// Characterization of the safe state per error class that had no test (#24 aim 6, step 1 of specs/plans/2026-11-02-reference-
// implementation-issue-24.md; the table is specs/design/monetcommon-safe-states.md). These tests pin what FB_MonetTelescopeControl
// does today on mock axes, with the line of the behaviour in a comment; they are not a specification. A test whose name ends in
// _Current pins a behaviour that differs from the target of the table (decision D4) and is flipped by the fix (step 7). The
// Roof_Request_* tests and No_Roof_Request_On_Focus_Error specify bCloseRoofRequest (step 7 PR 1, D9; no clock, no power-on). Every test
// owns a rig and runs over many PLC cycles (VAR_INST of the method, one Scan() per cycle). Failed checks are also noted in
// GVL_Diag.sFailures (printed by Run-Tests.ps1).
FUNCTION_BLOCK MonetSafeState_Tests EXTENDS TcUnit.FB_TestSuite
VAR
END_VAR

Hydraulics_Error_While_Tracking_Ramps_Then_Parks_In_Place();
Hydraulics_Pressure_Loss_While_Tracking_Parks_In_Place_Without_Ramp();
Cover_Error_At_PowerOn_Fails_And_Stays_Parked();
Cover_Error_During_Park_Ends_The_Park_Without_Closed();
Cover_Error_While_Tracking_Drives_To_Park();
Estop_During_Slew_Locks_Then_Parks_In_Place_After_The_Release();
Safety_Error_While_Tracking_Locks_Then_Parks_In_Place_When_It_Clears();
Power_Failure_During_Goto_Ramps_Then_Parks_In_Place();
Power_Failure_With_Pressure_Loss_Parks_In_Place_Without_Ramp();
Goto_Times_Out_Ramps_Then_Drives_To_Park();
Home_Times_Out_Ramps_Then_Drives_To_Park();
Clock_Invalid_Slew_Input_Is_Rejected();
Watchdog_Parks_And_Closes_The_Roof_In_One_Scan();
Invalid_Motion_Config_Is_Software_Error_32();
Roof_Request_On_Axis_Errors();
Roof_Request_On_Hydraulics_Error();
Roof_Request_On_Estop();
Roof_Request_On_Safety_Error();
Roof_Request_On_Power_Failure();
No_Roof_Request_On_Focus_Error();

// #24 step 7 PR 3 (D8, row hydraulics error; until 0.13.0 Hydraulics_Error_While_Tracking_Keeps_Tracking_Current): a hydraulics error
// with the pressure still there (brake open) is a telescope error (bHwError) and ramps first: in the scan of the error bStop is set
// (stop transaction, #96) and the axes stay enabled; every axis is sent its MC_Stop while still enabled (no 0x4257). After the stop
// has settled the emergency park queued behind it (bParkAfterStop) parks in place: axes disabled, brake closed, covers closed,
// hydraulics off, bIsParked and bParkedInPlace; READY_STATE -1.0 and bCloseRoofRequest while the error stays.
METHOD PRIVATE Hydraulics_Error_While_Tracking_Ramps_Then_Parks_In_Place
VAR_INST
	rig			: FB_MonetRig;
	nStep		: INT;
	nCycles		: UINT;
	nTracking	: UINT;
	sTest		: STRING(80);
	nEl0		: UINT;	// stop edges per axis before the error
	nAz0		: UINT;
	nDr0		: UINT;
	nExt0		: UINT;	// 0x4257 rejections of the three axes before the error
	nEdgesLast	: UINT;
	nEdgesNow	: UINT;
	nDisable0	: UINT;
	bSawStop	: BOOL;
	bStopOnDisabled	: BOOL;	// a stop edge came in a scan in which an axis was already disabled
END_VAR
TEST('Hydraulics_Error_While_Tracking_Ramps_Then_Parks_In_Place');
sTest := 'Hydraulics_Error_While_Tracking_Ramps_Then_Parks_In_Place: ';
IF nStep >= 90 THEN
	RETURN;
END_IF
rig.Scan();
nCycles := nCycles + 1;
CASE nStep OF
0:	// wait for the clock, then power on
	IF rig.ClockValid THEN
		rig.fbTel.Init();
		nStep := 10;
		nCycles := 0;
	ELSIF nCycles > 2000 THEN
		AssertTrue(Condition := FALSE, Message := 'the astronomical clock never became valid');
		F_Note(bFailed := TRUE, sText := CONCAT(sTest, 'the astronomical clock never became valid'));
		nStep := 99;
		TEST_FINISHED();
	END_IF
10:	// online: track a circumpolar target (always above the horizon, any RA)
	IF rig.Online THEN
		rig.fbTel.Track(fRightAscension := 0.0, fDeclination := -85.0);
		nStep := 20;
		nCycles := 0;
	ELSIF nCycles > 1500 THEN
		AssertTrue(Condition := FALSE, Message := 'the mock telescope did not reach READY_STATE 1.0');
		F_Note(bFailed := TRUE, sText := CONCAT(sTest, 'the mock telescope did not reach READY_STATE 1.0'));
		nStep := 99;
		TEST_FINISHED();
	END_IF
20:	// wait until all three axes have tracked for a few scans, then the hydraulics report an error (pressure still there)
	IF rig.fbAzim.Tracking AND rig.fbElev.Tracking AND rig.fbDero.Tracking THEN
		nTracking := nTracking + 1;
	ELSE
		nTracking := 0;
	END_IF
	IF nTracking >= 5 THEN
		nEl0 := rig.fbElev.nStopEdges;
		nAz0 := rig.fbAzim.nStopEdges;
		nDr0 := rig.fbDero.nStopEdges;
		nEdgesLast := nEl0 + nAz0 + nDr0;
		nExt0 := rig.fbElev.nExtErrors + rig.fbAzim.nExtErrors + rig.fbDero.nExtErrors;
		nDisable0 := rig.fbBrakeHyd.nDisableCalls;
		rig.fbBrakeHyd.InjectError();
		nStep := 30;
		nCycles := 0;
	ELSIF nCycles > 800 THEN
		AssertTrue(Condition := FALSE, Message := 'the telescope did not start tracking');
		F_Note(bFailed := TRUE, sText := CONCAT(sTest, 'the telescope did not start tracking'));
		nStep := 99;
		TEST_FINISHED();
	END_IF
30:	// ramp, then the park in place
	bSawStop := bSawStop OR rig.fbTel.bStopActive;
	nEdgesNow := rig.fbElev.nStopEdges + rig.fbAzim.nStopEdges + rig.fbDero.nStopEdges;
	IF nEdgesNow > nEdgesLast AND NOT (rig.fbElev.bEnable AND rig.fbAzim.bEnable AND rig.fbDero.bEnable) THEN
		bStopOnDisabled := TRUE;
	END_IF
	nEdgesLast := nEdgesNow;
	IF nCycles = 1 THEN	// the scan that saw the error
		AssertTrue(Condition := rig.fbTel.bStopActive AND rig.fbTel.bError, Message := 'the error stops the axes in its scan (bStop) and is a telescope error');
		F_Note(bFailed := NOT (rig.fbTel.bStopActive AND rig.fbTel.bError), sText := CONCAT(sTest, 'the error stops the axes in its scan (bStop) and is a telescope error'));
		AssertTrue(Condition := rig.fbElev.bEnable AND rig.fbAzim.bEnable AND rig.fbDero.bEnable, Message := 'the axes stay enabled for the ramp');
		F_Note(bFailed := NOT (rig.fbElev.bEnable AND rig.fbAzim.bEnable AND rig.fbDero.bEnable), sText := CONCAT(sTest, 'the axes stay enabled for the ramp'));
	END_IF
	IF rig.fbTel.bIsParked AND nCycles > 5 THEN
		AssertTrue(Condition := bSawStop, Message := 'the hydraulics error ramped (bStop)');
		F_Note(bFailed := NOT (bSawStop), sText := CONCAT(sTest, 'the hydraulics error ramped (bStop)'));
		AssertTrue(Condition := rig.fbElev.nStopEdges > nEl0 AND rig.fbAzim.nStopEdges > nAz0 AND rig.fbDero.nStopEdges > nDr0, Message := 'every axis was sent its MC_Stop');
		F_Note(bFailed := NOT (rig.fbElev.nStopEdges > nEl0 AND rig.fbAzim.nStopEdges > nAz0 AND rig.fbDero.nStopEdges > nDr0), sText := CONCAT(sTest, 'every axis was sent its MC_Stop'));
		AssertFalse(Condition := bStopOnDisabled, Message := 'the stops came before the disable');
		F_Note(bFailed := (bStopOnDisabled), sText := CONCAT(sTest, 'the stops came before the disable'));
		AssertTrue(Condition := rig.fbElev.nExtErrors + rig.fbAzim.nExtErrors + rig.fbDero.nExtErrors = nExt0, Message := 'no stop met the setpoint generator (0x4257)');
		F_Note(bFailed := NOT (rig.fbElev.nExtErrors + rig.fbAzim.nExtErrors + rig.fbDero.nExtErrors = nExt0), sText := CONCAT(sTest, 'no stop met the setpoint generator (0x4257)'));
		AssertTrue(Condition := rig.fbTel.bParkedInPlace AND NOT rig.fbTel.bParkActive, Message := 'the park ended in place');
		F_Note(bFailed := NOT (rig.fbTel.bParkedInPlace AND NOT rig.fbTel.bParkActive), sText := CONCAT(sTest, 'the park ended in place'));
		AssertFalse(Condition := rig.fbElev.bEnable OR rig.fbAzim.bEnable OR rig.fbDero.bEnable, Message := 'all three axes are disabled');
		F_Note(bFailed := (rig.fbElev.bEnable OR rig.fbAzim.bEnable OR rig.fbDero.bEnable), sText := CONCAT(sTest, 'all three axes are disabled'));
		AssertFalse(Condition := rig.fbBrakeHyd.BrakeOpen, Message := 'the brake is closed');
		F_Note(bFailed := (rig.fbBrakeHyd.BrakeOpen), sText := CONCAT(sTest, 'the brake is closed'));
		AssertTrue(Condition := rig.fbCovers.bClosed AND rig.fbCovers.nCloseCalls >= 1, Message := 'the covers are closed');
		F_Note(bFailed := NOT (rig.fbCovers.bClosed AND rig.fbCovers.nCloseCalls >= 1), sText := CONCAT(sTest, 'the covers are closed'));
		AssertTrue(Condition := rig.fbBrakeHyd.nDisableCalls > nDisable0, Message := 'the hydraulics are switched off');
		F_Note(bFailed := NOT (rig.fbBrakeHyd.nDisableCalls > nDisable0), sText := CONCAT(sTest, 'the hydraulics are switched off'));
		AssertFalse(Condition := rig.fbTel.bTrackActive OR rig.fbAzim.Tracking OR rig.fbElev.Tracking OR rig.fbDero.Tracking, Message := 'nothing tracks any more');
		F_Note(bFailed := (rig.fbTel.bTrackActive OR rig.fbAzim.Tracking OR rig.fbElev.Tracking OR rig.fbDero.Tracking), sText := CONCAT(sTest, 'nothing tracks any more'));
		AssertTrue(Condition := rig.fbTel.bError AND rig.fbTel.ReadyState = -1.0, Message := 'the error stays, READY_STATE -1.0');
		F_Note(bFailed := NOT (rig.fbTel.bError AND rig.fbTel.ReadyState = -1.0), sText := CONCAT(sTest, 'the error stays, READY_STATE -1.0'));
		AssertTrue(Condition := rig.fbTel.bCloseRoofRequest, Message := 'the roof close is requested');
		F_Note(bFailed := NOT (rig.fbTel.bCloseRoofRequest), sText := CONCAT(sTest, 'the roof close is requested'));
		nStep := 99;
		TEST_FINISHED();
	ELSIF nCycles > 800 THEN
		AssertTrue(Condition := FALSE, Message := 'the telescope did not park after the ramp');
		F_Note(bFailed := TRUE, sText := CONCAT(sTest, 'the telescope did not park after the ramp'));
		nStep := 99;
		TEST_FINISHED();
	END_IF
END_CASE
END_METHOD

// #24 step 7 PR 3 (D8, row hydraulics error): a hydraulics error with the oil pressure already gone (mock InjectPressureLoss: the
// brake is locked) cannot ramp, the brake lock is the stop: the axes are disabled in the scan of the error, as for an axis error,
// no MC_Stop is sent, and the emergency park parks in place (covers closed, hydraulics off, bIsParked, bParkedInPlace).
METHOD PRIVATE Hydraulics_Pressure_Loss_While_Tracking_Parks_In_Place_Without_Ramp
VAR_INST
	rig			: FB_MonetRig;
	nStep		: INT;
	nCycles		: UINT;
	nTracking	: UINT;
	sTest		: STRING(80);
	nEdges0		: UINT;	// stop edges of the three axes before the error
	nDisable0	: UINT;
	bSawStop	: BOOL;
END_VAR
TEST('Hydraulics_Pressure_Loss_While_Tracking_Parks_In_Place_Without_Ramp');
sTest := 'Hydraulics_Pressure_Loss_While_Tracking_Parks_In_Place_Without_Ramp: ';
IF nStep >= 90 THEN
	RETURN;
END_IF
rig.Scan();
nCycles := nCycles + 1;
CASE nStep OF
0:	// wait for the clock, then power on
	IF rig.ClockValid THEN
		rig.fbTel.Init();
		nStep := 10;
		nCycles := 0;
	ELSIF nCycles > 2000 THEN
		AssertTrue(Condition := FALSE, Message := 'the astronomical clock never became valid');
		F_Note(bFailed := TRUE, sText := CONCAT(sTest, 'the astronomical clock never became valid'));
		nStep := 99;
		TEST_FINISHED();
	END_IF
10:	// online: track a circumpolar target
	IF rig.Online THEN
		rig.fbTel.Track(fRightAscension := 0.0, fDeclination := -85.0);
		nStep := 20;
		nCycles := 0;
	ELSIF nCycles > 1500 THEN
		AssertTrue(Condition := FALSE, Message := 'the mock telescope did not reach READY_STATE 1.0');
		F_Note(bFailed := TRUE, sText := CONCAT(sTest, 'the mock telescope did not reach READY_STATE 1.0'));
		nStep := 99;
		TEST_FINISHED();
	END_IF
20:	// tracking: the hydraulics fail and the pressure is gone at once (the brake locks)
	IF rig.fbAzim.Tracking AND rig.fbElev.Tracking AND rig.fbDero.Tracking THEN
		nTracking := nTracking + 1;
	ELSE
		nTracking := 0;
	END_IF
	IF nTracking >= 5 THEN
		nEdges0 := rig.fbElev.nStopEdges + rig.fbAzim.nStopEdges + rig.fbDero.nStopEdges;
		nDisable0 := rig.fbBrakeHyd.nDisableCalls;
		rig.fbBrakeHyd.InjectPressureLoss();
		nStep := 30;
		nCycles := 0;
	ELSIF nCycles > 800 THEN
		AssertTrue(Condition := FALSE, Message := 'the telescope did not start tracking');
		F_Note(bFailed := TRUE, sText := CONCAT(sTest, 'the telescope did not start tracking'));
		nStep := 99;
		TEST_FINISHED();
	END_IF
30:
	bSawStop := bSawStop OR rig.fbTel.bStopActive;
	IF nCycles = 1 THEN	// the scan that saw the error
		AssertFalse(Condition := rig.fbElev.bEnable OR rig.fbAzim.bEnable OR rig.fbDero.bEnable, Message := 'the lock is the stop: disabled in the scan of the error');
		F_Note(bFailed := (rig.fbElev.bEnable OR rig.fbAzim.bEnable OR rig.fbDero.bEnable), sText := CONCAT(sTest, 'the lock is the stop: disabled in the scan of the error'));
	END_IF
	IF rig.fbTel.bIsParked AND nCycles > 5 THEN
		AssertFalse(Condition := bSawStop, Message := 'no ramp (bStop never set)');
		F_Note(bFailed := (bSawStop), sText := CONCAT(sTest, 'no ramp (bStop never set)'));
		AssertTrue(Condition := rig.fbElev.nStopEdges + rig.fbAzim.nStopEdges + rig.fbDero.nStopEdges = nEdges0, Message := 'no MC_Stop was sent');
		F_Note(bFailed := NOT (rig.fbElev.nStopEdges + rig.fbAzim.nStopEdges + rig.fbDero.nStopEdges = nEdges0), sText := CONCAT(sTest, 'no MC_Stop was sent'));
		AssertTrue(Condition := rig.fbTel.bParkedInPlace AND NOT rig.fbTel.bParkActive, Message := 'the park ended in place');
		F_Note(bFailed := NOT (rig.fbTel.bParkedInPlace AND NOT rig.fbTel.bParkActive), sText := CONCAT(sTest, 'the park ended in place'));
		AssertFalse(Condition := rig.fbBrakeHyd.BrakeOpen, Message := 'the brake is locked');
		F_Note(bFailed := (rig.fbBrakeHyd.BrakeOpen), sText := CONCAT(sTest, 'the brake is locked'));
		AssertTrue(Condition := rig.fbCovers.bClosed AND rig.fbCovers.nCloseCalls >= 1, Message := 'the covers are closed');
		F_Note(bFailed := NOT (rig.fbCovers.bClosed AND rig.fbCovers.nCloseCalls >= 1), sText := CONCAT(sTest, 'the covers are closed'));
		AssertTrue(Condition := rig.fbBrakeHyd.nDisableCalls > nDisable0, Message := 'the hydraulics are switched off');
		F_Note(bFailed := NOT (rig.fbBrakeHyd.nDisableCalls > nDisable0), sText := CONCAT(sTest, 'the hydraulics are switched off'));
		AssertTrue(Condition := rig.fbTel.bError AND rig.fbTel.ReadyState = -1.0, Message := 'the error stays, READY_STATE -1.0');
		F_Note(bFailed := NOT (rig.fbTel.bError AND rig.fbTel.ReadyState = -1.0), sText := CONCAT(sTest, 'the error stays, READY_STATE -1.0'));
		AssertTrue(Condition := rig.fbTel.bCloseRoofRequest, Message := 'the roof close is requested');
		F_Note(bFailed := NOT (rig.fbTel.bCloseRoofRequest), sText := CONCAT(sTest, 'the roof close is requested'));
		nStep := 99;
		TEST_FINISHED();
	ELSIF nCycles > 800 THEN
		AssertTrue(Condition := FALSE, Message := 'the emergency park did not finish');
		F_Note(bFailed := TRUE, sText := CONCAT(sTest, 'the emergency park did not finish'));
		nStep := 99;
		TEST_FINISHED();
	END_IF
END_CASE
END_METHOD

// #24 step 7 PR 4 (row cover error; until 0.13.x Cover_Error_At_PowerOn_Waits_In_Stage_0_Current, where the power-on waited in
// stage 0 for fbCovers.Opened until the 12 h command timeout, with bIsParked already FALSE). A cover error on a parked telescope
// starts no park. A power-on with the cover error fails in its first scan, before the cover command of stage 0 (_PowerOn checks,
// bPowerFailure): nothing opens, no axis is enabled, the telescope stays parked, READY_STATE -1.0, no telescope error, no roof
// close request (D9). Reset path: the cover reset (HalfBROT Reset(), MAIN reset button), then power=1 goes online.
METHOD PRIVATE Cover_Error_At_PowerOn_Fails_And_Stays_Parked
VAR_INST
	rig			: FB_MonetRig;
	nStep		: INT;
	nCycles		: UINT;
	sTest		: STRING(80);
END_VAR
TEST('Cover_Error_At_PowerOn_Fails_And_Stays_Parked');
sTest := 'Cover_Error_At_PowerOn_Fails_And_Stays_Parked: ';
IF nStep >= 90 THEN
	RETURN;
END_IF
rig.Scan();
nCycles := nCycles + 1;
CASE nStep OF
0:	// wait for the clock; the covers of the parked telescope report an error
	IF rig.ClockValid THEN
		rig.fbCovers.InjectError();
		nStep := 5;
		nCycles := 0;
	ELSIF nCycles > 2000 THEN
		AssertTrue(Condition := FALSE, Message := 'the astronomical clock never became valid');
		F_Note(bFailed := TRUE, sText := CONCAT(sTest, 'the astronomical clock never became valid'));
		nStep := 99;
		TEST_FINISHED();
	END_IF
5:	// parked: nothing happens; then power on
	IF nCycles >= 10 THEN
		AssertTrue(Condition := rig.fbTel.bIsParked AND NOT rig.fbTel.bParkActive AND NOT rig.fbTel.bError, Message := 'a cover error on a parked telescope starts no park and is no telescope error');
		F_Note(bFailed := NOT (rig.fbTel.bIsParked AND NOT rig.fbTel.bParkActive AND NOT rig.fbTel.bError), sText := CONCAT(sTest, 'a cover error on a parked telescope starts no park and is no telescope error'));
		rig.fbTel.Init();
		nStep := 10;
		nCycles := 0;
	END_IF
10:	// the power-on fails in its first scan
	IF nCycles >= 10 THEN
		AssertFalse(Condition := rig.fbTel.bPowerActive OR rig.fbTel.fbStartup.Initializing, Message := 'the power-on is over');
		F_Note(bFailed := (rig.fbTel.bPowerActive OR rig.fbTel.fbStartup.Initializing), sText := CONCAT(sTest, 'the power-on is over'));
		AssertTrue(Condition := rig.fbTel.bPowerFailure AND rig.fbTel.ReadyState = -1.0, Message := 'power-on failure, READY_STATE -1.0');
		F_Note(bFailed := NOT (rig.fbTel.bPowerFailure AND rig.fbTel.ReadyState = -1.0), sText := CONCAT(sTest, 'power-on failure, READY_STATE -1.0'));
		AssertTrue(Condition := rig.fbCovers.nOpenCalls = 0 AND NOT rig.fbCovers.bOpened, Message := 'the covers were not commanded');
		F_Note(bFailed := NOT (rig.fbCovers.nOpenCalls = 0 AND NOT rig.fbCovers.bOpened), sText := CONCAT(sTest, 'the covers were not commanded'));
		AssertFalse(Condition := rig.fbElev.bEnable OR rig.fbAzim.bEnable OR rig.fbDero.bEnable, Message := 'no axis was enabled');
		F_Note(bFailed := (rig.fbElev.bEnable OR rig.fbAzim.bEnable OR rig.fbDero.bEnable), sText := CONCAT(sTest, 'no axis was enabled'));
		AssertTrue(Condition := rig.fbTel.bIsParked, Message := 'the telescope stays parked');
		F_Note(bFailed := NOT (rig.fbTel.bIsParked), sText := CONCAT(sTest, 'the telescope stays parked'));
		AssertFalse(Condition := rig.fbTel.bError, Message := 'a cover error is not a telescope error');
		F_Note(bFailed := (rig.fbTel.bError), sText := CONCAT(sTest, 'a cover error is not a telescope error'));
		AssertFalse(Condition := rig.fbTel.bCloseRoofRequest, Message := 'no roof close request for a cover error');
		F_Note(bFailed := (rig.fbTel.bCloseRoofRequest), sText := CONCAT(sTest, 'no roof close request for a cover error'));
		rig.fbCovers.Reset();	// MAIN reset button
		nStep := 20;
		nCycles := 0;
	END_IF
20:
	IF nCycles >= 3 THEN
		rig.fbTel.Init();
		nStep := 30;
		nCycles := 0;
	END_IF
30:	// power=1 after the cover reset: online
	IF rig.Online THEN
		AssertTrue(Condition := rig.fbCovers.bOpened AND NOT rig.fbTel.bPowerFailure, Message := 'online after the cover reset and power=1');
		F_Note(bFailed := NOT (rig.fbCovers.bOpened AND NOT rig.fbTel.bPowerFailure), sText := CONCAT(sTest, 'online after the cover reset and power=1'));
		nStep := 99;
		TEST_FINISHED();
	ELSIF nCycles > 1500 THEN
		AssertTrue(Condition := FALSE, Message := 'not online after the cover reset and power=1');
		F_Note(bFailed := TRUE, sText := CONCAT(sTest, 'not online after the cover reset and power=1'));
		nStep := 99;
		TEST_FINISHED();
	END_IF
END_CASE
END_METHOD

// #24 step 7 PR 4 (row cover error; until 0.13.x Cover_Error_Holds_The_Park_Before_Parked_Current, where the park waited in stage
// secure for fbCovers.Closed for ever: bPark held, READY_STATE 0.3, never bIsParked). A cover error during the drive to the park
// position: the park goes on (no telescope error, the drives are controllable), reaches the park position, disables the axes, the
// brake closes, the hydraulics go off, and the park ends without Closed: bIsParked, not in place, software error 16#21 (READY_STATE
// -1.0), no roof close request (D9).
METHOD PRIVATE Cover_Error_During_Park_Ends_The_Park_Without_Closed
VAR_INST
	rig			: FB_MonetRig;
	nStep		: INT;
	nCycles		: UINT;
	sTest		: STRING(80);
	nDisable0	: UINT;
	bSawError	: BOOL;	// bError before the park ended
END_VAR
TEST('Cover_Error_During_Park_Ends_The_Park_Without_Closed');
sTest := 'Cover_Error_During_Park_Ends_The_Park_Without_Closed: ';
IF nStep >= 90 THEN
	RETURN;
END_IF
rig.Scan();
nCycles := nCycles + 1;
CASE nStep OF
0:	// wait for the clock, then power on
	IF rig.ClockValid THEN
		rig.fbTel.Init();
		nStep := 10;
		nCycles := 0;
	ELSIF nCycles > 2000 THEN
		AssertTrue(Condition := FALSE, Message := 'the astronomical clock never became valid');
		F_Note(bFailed := TRUE, sText := CONCAT(sTest, 'the astronomical clock never became valid'));
		nStep := 99;
		TEST_FINISHED();
	END_IF
10:	// online: slow axes, park
	IF rig.Online THEN
		rig.SetMoveScans(nScans := 300);
		nDisable0 := rig.fbBrakeHyd.nDisableCalls;
		rig.fbTel.Park();
		nStep := 20;
		nCycles := 0;
	ELSIF nCycles > 1500 THEN
		AssertTrue(Condition := FALSE, Message := 'the mock telescope did not reach READY_STATE 1.0');
		F_Note(bFailed := TRUE, sText := CONCAT(sTest, 'the mock telescope did not reach READY_STATE 1.0'));
		nStep := 99;
		TEST_FINISHED();
	END_IF
20:	// the park drives: the covers report an error
	IF rig.fbElev.MoveAxis AND rig.fbAzim.MoveAxis AND rig.fbDero.MoveAxis AND nCycles > 5 THEN
		rig.fbCovers.InjectError();
		nStep := 30;
		nCycles := 0;
	ELSIF nCycles > 300 THEN
		AssertTrue(Condition := FALSE, Message := 'the park did not start the axis moves');
		F_Note(bFailed := TRUE, sText := CONCAT(sTest, 'the park did not start the axis moves'));
		nStep := 99;
		TEST_FINISHED();
	END_IF
30:	// the park goes on and ends
	IF rig.fbTel.bIsParked THEN
		AssertFalse(Condition := bSawError, Message := 'no telescope error during the drive');
		F_Note(bFailed := (bSawError), sText := CONCAT(sTest, 'no telescope error during the drive'));
		AssertFalse(Condition := rig.fbTel.bParkActive OR rig.fbTel.bParkedInPlace, Message := 'the park is over, not in place');
		F_Note(bFailed := (rig.fbTel.bParkActive OR rig.fbTel.bParkedInPlace), sText := CONCAT(sTest, 'the park is over, not in place'));
		AssertTrue(Condition := ABS(rig.fbElev.fActualPosition - 60.0) < 0.001 AND ABS(rig.fbAzim.fActualPosition - 175.0) < 0.001, Message := 'at the park position');
		F_Note(bFailed := NOT (ABS(rig.fbElev.fActualPosition - 60.0) < 0.001 AND ABS(rig.fbAzim.fActualPosition - 175.0) < 0.001), sText := CONCAT(sTest, 'at the park position'));
		AssertFalse(Condition := rig.fbElev.bEnable OR rig.fbAzim.bEnable OR rig.fbDero.bEnable, Message := 'all three axes are disabled');
		F_Note(bFailed := (rig.fbElev.bEnable OR rig.fbAzim.bEnable OR rig.fbDero.bEnable), sText := CONCAT(sTest, 'all three axes are disabled'));
		AssertFalse(Condition := rig.fbBrakeHyd.BrakeOpen, Message := 'the brake is closed');
		F_Note(bFailed := (rig.fbBrakeHyd.BrakeOpen), sText := CONCAT(sTest, 'the brake is closed'));
		AssertTrue(Condition := rig.fbBrakeHyd.nDisableCalls > nDisable0, Message := 'the hydraulics are switched off');
		F_Note(bFailed := NOT (rig.fbBrakeHyd.nDisableCalls > nDisable0), sText := CONCAT(sTest, 'the hydraulics are switched off'));
		AssertTrue(Condition := rig.fbCovers.nCloseCalls >= 1 AND NOT rig.fbCovers.bClosed, Message := 'the covers were commanded closed and did not move');
		F_Note(bFailed := NOT (rig.fbCovers.nCloseCalls >= 1 AND NOT rig.fbCovers.bClosed), sText := CONCAT(sTest, 'the covers were commanded closed and did not move'));
		AssertTrue(Condition := rig.fbTel.bError AND rig.fbTel.nErrorID = 16#21 AND rig.fbTel.ReadyState = -1.0, Message := 'software error 16#21, READY_STATE -1.0');
		F_Note(bFailed := NOT (rig.fbTel.bError AND rig.fbTel.nErrorID = 16#21 AND rig.fbTel.ReadyState = -1.0), sText := CONCAT(sTest, 'software error 16#21, READY_STATE -1.0'));
		AssertFalse(Condition := rig.fbTel.bCloseRoofRequest, Message := 'no roof close request for a cover error');
		F_Note(bFailed := (rig.fbTel.bCloseRoofRequest), sText := CONCAT(sTest, 'no roof close request for a cover error'));
		nStep := 99;
		TEST_FINISHED();
	ELSIF nCycles > 1500 THEN
		AssertTrue(Condition := FALSE, Message := 'the park did not end (it waits for the covers)');
		F_Note(bFailed := TRUE, sText := CONCAT(sTest, 'the park did not end (it waits for the covers)'));
		nStep := 99;
		TEST_FINISHED();
	END_IF
	bSawError := bSawError OR rig.fbTel.bError;	// after the check: 16#21 is raised in the scan that sets bIsParked
END_CASE
END_METHOD

// #24 step 7 PR 4 (row cover error, target "ramp; drive to park"): a cover error while tracking is no telescope error (the drives are
// controllable) and starts a normal park in its scan (Park(), the routing of an external park: the track is dropped, the axes stay
// enabled and drive to the park position). The park ends without Closed: bIsParked, not in place, hydraulics off, software error
// 16#21, no roof close request (D9).
METHOD PRIVATE Cover_Error_While_Tracking_Drives_To_Park
VAR_INST
	rig			: FB_MonetRig;
	nStep		: INT;
	nCycles		: UINT;
	nTracking	: UINT;
	sTest		: STRING(80);
	nDisable0	: UINT;
END_VAR
TEST('Cover_Error_While_Tracking_Drives_To_Park');
sTest := 'Cover_Error_While_Tracking_Drives_To_Park: ';
IF nStep >= 90 THEN
	RETURN;
END_IF
rig.Scan();
nCycles := nCycles + 1;
CASE nStep OF
0:	// wait for the clock, then power on
	IF rig.ClockValid THEN
		rig.fbTel.Init();
		nStep := 10;
		nCycles := 0;
	ELSIF nCycles > 2000 THEN
		AssertTrue(Condition := FALSE, Message := 'the astronomical clock never became valid');
		F_Note(bFailed := TRUE, sText := CONCAT(sTest, 'the astronomical clock never became valid'));
		nStep := 99;
		TEST_FINISHED();
	END_IF
10:	// online: track a circumpolar target
	IF rig.Online THEN
		rig.fbTel.Track(fRightAscension := 0.0, fDeclination := -85.0);
		nStep := 20;
		nCycles := 0;
	ELSIF nCycles > 1500 THEN
		AssertTrue(Condition := FALSE, Message := 'the mock telescope did not reach READY_STATE 1.0');
		F_Note(bFailed := TRUE, sText := CONCAT(sTest, 'the mock telescope did not reach READY_STATE 1.0'));
		nStep := 99;
		TEST_FINISHED();
	END_IF
20:	// tracking: the covers report an error
	IF rig.fbAzim.Tracking AND rig.fbElev.Tracking AND rig.fbDero.Tracking THEN
		nTracking := nTracking + 1;
	ELSE
		nTracking := 0;
	END_IF
	IF nTracking >= 5 THEN
		nDisable0 := rig.fbBrakeHyd.nDisableCalls;
		rig.fbCovers.InjectError();
		nStep := 30;
		nCycles := 0;
	ELSIF nCycles > 800 THEN
		AssertTrue(Condition := FALSE, Message := 'the telescope did not start tracking');
		F_Note(bFailed := TRUE, sText := CONCAT(sTest, 'the telescope did not start tracking'));
		nStep := 99;
		TEST_FINISHED();
	END_IF
30:
	IF nCycles = 1 THEN	// the scan that saw the error
		AssertTrue(Condition := rig.fbTel.bParkActive AND NOT rig.fbTel.bTrackActive, Message := 'the park is requested in the scan of the error, the track is dropped');
		F_Note(bFailed := NOT (rig.fbTel.bParkActive AND NOT rig.fbTel.bTrackActive), sText := CONCAT(sTest, 'the park is requested in the scan of the error, the track is dropped'));
		AssertTrue(Condition := NOT rig.fbTel.bError AND rig.fbElev.bEnable AND rig.fbAzim.bEnable AND rig.fbDero.bEnable, Message := 'no telescope error, the axes stay enabled');
		F_Note(bFailed := NOT (NOT rig.fbTel.bError AND rig.fbElev.bEnable AND rig.fbAzim.bEnable AND rig.fbDero.bEnable), sText := CONCAT(sTest, 'no telescope error, the axes stay enabled'));
	END_IF
	IF rig.fbTel.bIsParked AND nCycles > 5 THEN
		AssertFalse(Condition := rig.fbTel.bParkActive OR rig.fbTel.bParkedInPlace, Message := 'the park is over, not in place');
		F_Note(bFailed := (rig.fbTel.bParkActive OR rig.fbTel.bParkedInPlace), sText := CONCAT(sTest, 'the park is over, not in place'));
		AssertTrue(Condition := ABS(rig.fbElev.fActualPosition - 60.0) < 0.001 AND ABS(rig.fbAzim.fActualPosition - 175.0) < 0.001, Message := 'at the park position');
		F_Note(bFailed := NOT (ABS(rig.fbElev.fActualPosition - 60.0) < 0.001 AND ABS(rig.fbAzim.fActualPosition - 175.0) < 0.001), sText := CONCAT(sTest, 'at the park position'));
		AssertFalse(Condition := rig.fbTel.bTrackActive OR rig.fbAzim.Tracking OR rig.fbElev.Tracking OR rig.fbDero.Tracking, Message := 'nothing tracks any more');
		F_Note(bFailed := (rig.fbTel.bTrackActive OR rig.fbAzim.Tracking OR rig.fbElev.Tracking OR rig.fbDero.Tracking), sText := CONCAT(sTest, 'nothing tracks any more'));
		AssertFalse(Condition := rig.fbElev.bEnable OR rig.fbAzim.bEnable OR rig.fbDero.bEnable OR rig.fbBrakeHyd.BrakeOpen, Message := 'axes disabled, brake closed');
		F_Note(bFailed := (rig.fbElev.bEnable OR rig.fbAzim.bEnable OR rig.fbDero.bEnable OR rig.fbBrakeHyd.BrakeOpen), sText := CONCAT(sTest, 'axes disabled, brake closed'));
		AssertTrue(Condition := rig.fbBrakeHyd.nDisableCalls > nDisable0, Message := 'the hydraulics are switched off');
		F_Note(bFailed := NOT (rig.fbBrakeHyd.nDisableCalls > nDisable0), sText := CONCAT(sTest, 'the hydraulics are switched off'));
		AssertFalse(Condition := rig.fbCovers.bClosed, Message := 'the covers did not move');
		F_Note(bFailed := (rig.fbCovers.bClosed), sText := CONCAT(sTest, 'the covers did not move'));
		AssertTrue(Condition := rig.fbTel.nErrorID = 16#21 AND rig.fbTel.ReadyState = -1.0, Message := 'software error 16#21, READY_STATE -1.0');
		F_Note(bFailed := NOT (rig.fbTel.nErrorID = 16#21 AND rig.fbTel.ReadyState = -1.0), sText := CONCAT(sTest, 'software error 16#21, READY_STATE -1.0'));
		AssertFalse(Condition := rig.fbTel.bCloseRoofRequest, Message := 'no roof close request for a cover error');
		F_Note(bFailed := (rig.fbTel.bCloseRoofRequest), sText := CONCAT(sTest, 'no roof close request for a cover error'));
		nStep := 99;
		TEST_FINISHED();
	ELSIF nCycles > 1500 THEN
		AssertTrue(Condition := FALSE, Message := 'the park did not end');
		F_Note(bFailed := TRUE, sText := CONCAT(sTest, 'the park did not end'));
		nStep := 99;
		TEST_FINISHED();
	END_IF
END_CASE
END_METHOD

// #24 step 7 PR 6 (D8, row E-stop; until 0.13.0 Estop_During_Slew_Disables_The_Axes_Without_Park_Current): the E-stop under a slew
// is a lock stop: in its scan the three axes are disabled and the hydraulics switched off (the brake locks), no stop transaction
// (no bStop, no MC_Stop), the slew ends. During the E-stop nothing parks and the covers are not commanded (they may hang on the
// same circuit), also not after a reset (the MAIN reset button that starts the safety reset); READY_STATE -1.0, not bError. After
// the release (E-stop gone, safety reset done) the held park runs in place: covers closed, hydraulics off, bIsParked,
// bParkedInPlace; the roof request stays until a reset; then power=1 is online again. The mock axis keeps its move when it is
// disabled (STO is not modelled), so the test ends the mock move (SetMoveScans) before the release.
METHOD PRIVATE Estop_During_Slew_Locks_Then_Parks_In_Place_After_The_Release
VAR_INST
	rig			: FB_MonetRig;
	nStep		: INT;
	nCycles		: UINT;
	sTest		: STRING(80);
	nDisable0	: UINT;	// hydraulics-off writes before the E-stop
	nDisable1	: UINT;	// ... before the release
	nEdges0		: UINT;	// MC_Stop requests of the three axes before the E-stop
	bSawStop	: BOOL;
END_VAR
TEST('Estop_During_Slew_Locks_Then_Parks_In_Place_After_The_Release');
sTest := 'Estop_During_Slew_Locks_Then_Parks_In_Place_After_The_Release: ';
IF nStep >= 90 THEN
	RETURN;
END_IF
rig.Scan();
nCycles := nCycles + 1;
CASE nStep OF
0:	// wait for the clock, then power on
	IF rig.ClockValid THEN
		rig.fbTel.Init();
		nStep := 10;
		nCycles := 0;
	ELSIF nCycles > 2000 THEN
		AssertTrue(Condition := FALSE, Message := 'the astronomical clock never became valid');
		F_Note(bFailed := TRUE, sText := CONCAT(sTest, 'the astronomical clock never became valid'));
		nStep := 99;
		TEST_FINISHED();
	END_IF
10:	// online: slow axes, slew
	IF rig.Online THEN
		rig.SetMoveScans(nScans := 3000);
		rig.fbTel.Slew(fAzimuth := 180.0, fAltitude := 45.0);
		nStep := 20;
		nCycles := 0;
	ELSIF nCycles > 1500 THEN
		AssertTrue(Condition := FALSE, Message := 'the mock telescope did not reach READY_STATE 1.0');
		F_Note(bFailed := TRUE, sText := CONCAT(sTest, 'the mock telescope did not reach READY_STATE 1.0'));
		nStep := 99;
		TEST_FINISHED();
	END_IF
20:
	IF rig.fbElev.MoveAxis AND rig.fbAzim.MoveAxis AND rig.fbDero.MoveAxis THEN
		nStep := 30;
		nCycles := 0;
	ELSIF nCycles > 300 THEN
		AssertTrue(Condition := FALSE, Message := 'the slew did not start the axis moves');
		F_Note(bFailed := TRUE, sText := CONCAT(sTest, 'the slew did not start the axis moves'));
		nStep := 99;
		TEST_FINISHED();
	END_IF
30:	// the axes move: the E-stop is pressed
	IF nCycles >= 5 THEN
		nDisable0 := rig.fbBrakeHyd.nDisableCalls;
		nEdges0 := rig.fbElev.nStopEdges + rig.fbAzim.nStopEdges + rig.fbDero.nStopEdges;
		rig.SetEstop(TRUE);
		nStep := 40;
		nCycles := 0;
	END_IF
40:	// the lock is the stop; the park is held while the E-stop is pressed
	bSawStop := bSawStop OR rig.fbTel.bStopActive;
	IF nCycles = 1 THEN	// the scan that saw the E-stop
		AssertFalse(Condition := rig.fbElev.bEnable OR rig.fbAzim.bEnable OR rig.fbDero.bEnable, Message := 'the axes are disabled in the scan of the E-stop');
		F_Note(bFailed := (rig.fbElev.bEnable OR rig.fbAzim.bEnable OR rig.fbDero.bEnable), sText := CONCAT(sTest, 'the axes are disabled in the scan of the E-stop'));
		AssertTrue(Condition := rig.fbBrakeHyd.nDisableCalls > nDisable0, Message := 'the hydraulics go off in the scan of the E-stop');
		F_Note(bFailed := NOT (rig.fbBrakeHyd.nDisableCalls > nDisable0), sText := CONCAT(sTest, 'the hydraulics go off in the scan of the E-stop'));
		AssertTrue(Condition := rig.fbCovers.nStopCalls >= 1, Message := 'the covers get Stop() in the scan of the E-stop (not on the E-stop circuit)');
		F_Note(bFailed := NOT (rig.fbCovers.nStopCalls >= 1), sText := CONCAT(sTest, 'the covers get Stop() in the scan of the E-stop (not on the E-stop circuit)'));
	END_IF
	IF nCycles >= 60 THEN
		AssertFalse(Condition := rig.fbElev.bEnable OR rig.fbAzim.bEnable OR rig.fbDero.bEnable, Message := 'the three axes are disabled');
		F_Note(bFailed := (rig.fbElev.bEnable OR rig.fbAzim.bEnable OR rig.fbDero.bEnable), sText := CONCAT(sTest, 'the three axes are disabled'));
		AssertFalse(Condition := rig.fbBrakeHyd.BrakeOpen, Message := 'the brake is closed');
		F_Note(bFailed := (rig.fbBrakeHyd.BrakeOpen), sText := CONCAT(sTest, 'the brake is closed'));
		AssertFalse(Condition := bSawStop, Message := 'no ramp (bStop never set)');
		F_Note(bFailed := (bSawStop), sText := CONCAT(sTest, 'no ramp (bStop never set)'));
		AssertTrue(Condition := rig.fbElev.nStopEdges + rig.fbAzim.nStopEdges + rig.fbDero.nStopEdges = nEdges0, Message := 'no MC_Stop was sent');
		F_Note(bFailed := NOT (rig.fbElev.nStopEdges + rig.fbAzim.nStopEdges + rig.fbDero.nStopEdges = nEdges0), sText := CONCAT(sTest, 'no MC_Stop was sent'));
		AssertFalse(Condition := rig.fbTel.bSlewActive, Message := 'the slew has ended');
		F_Note(bFailed := (rig.fbTel.bSlewActive), sText := CONCAT(sTest, 'the slew has ended'));
		AssertFalse(Condition := rig.fbTel.bParkActive OR rig.fbTel.bIsParked, Message := 'no park during the E-stop');
		F_Note(bFailed := (rig.fbTel.bParkActive OR rig.fbTel.bIsParked), sText := CONCAT(sTest, 'no park during the E-stop'));
		AssertTrue(Condition := rig.fbCovers.nCloseCalls = 0, Message := 'the covers are not commanded during the E-stop');
		F_Note(bFailed := NOT (rig.fbCovers.nCloseCalls = 0), sText := CONCAT(sTest, 'the covers are not commanded during the E-stop'));
		AssertFalse(Condition := rig.fbTel.bError, Message := 'the E-stop is not bError');
		F_Note(bFailed := (rig.fbTel.bError), sText := CONCAT(sTest, 'the E-stop is not bError'));
		AssertTrue(Condition := rig.fbTel.ReadyState = -1.0, Message := 'READY_STATE is -1.0');
		F_Note(bFailed := NOT (rig.fbTel.ReadyState = -1.0), sText := CONCAT(sTest, 'READY_STATE is -1.0'));
		rig.SetMoveScans(nScans := 60);	// STO is not modelled: end the move the disabled mock axes still run
		rig.fbTel.Reset();	// the MAIN reset button during the E-stop (starts the safety reset)
		nStep := 50;
		nCycles := 0;
	END_IF
50:	// a reset during the E-stop does not start the park
	bSawStop := bSawStop OR rig.fbTel.bStopActive;
	IF nCycles >= 10 THEN
		AssertTrue(Condition := NOT (rig.fbTel.bParkActive OR rig.fbTel.bIsParked) AND rig.fbCovers.nCloseCalls = 0, Message := 'a reset during the E-stop does not start the park');
		F_Note(bFailed := NOT (NOT (rig.fbTel.bParkActive OR rig.fbTel.bIsParked) AND rig.fbCovers.nCloseCalls = 0), sText := CONCAT(sTest, 'a reset during the E-stop does not start the park'));
		nDisable1 := rig.fbBrakeHyd.nDisableCalls;
		rig.SetEstop(FALSE);	// released, safety reset done
		nStep := 60;
		nCycles := 0;
	END_IF
60:	// after the release: the park in place
	bSawStop := bSawStop OR rig.fbTel.bStopActive;
	IF rig.fbTel.bIsParked AND nCycles > 5 THEN
		AssertTrue(Condition := rig.fbTel.bParkedInPlace AND NOT rig.fbTel.bParkActive, Message := 'the park after the release ended in place');
		F_Note(bFailed := NOT (rig.fbTel.bParkedInPlace AND NOT rig.fbTel.bParkActive), sText := CONCAT(sTest, 'the park after the release ended in place'));
		AssertTrue(Condition := rig.fbCovers.bClosed AND rig.fbCovers.nCloseCalls >= 1, Message := 'the covers are closed after the release');
		F_Note(bFailed := NOT (rig.fbCovers.bClosed AND rig.fbCovers.nCloseCalls >= 1), sText := CONCAT(sTest, 'the covers are closed after the release'));
		AssertTrue(Condition := rig.fbBrakeHyd.nDisableCalls > nDisable1, Message := 'the park switches the hydraulics off');
		F_Note(bFailed := NOT (rig.fbBrakeHyd.nDisableCalls > nDisable1), sText := CONCAT(sTest, 'the park switches the hydraulics off'));
		AssertFalse(Condition := rig.fbElev.bEnable OR rig.fbAzim.bEnable OR rig.fbDero.bEnable OR rig.fbBrakeHyd.BrakeOpen, Message := 'axes disabled, brake closed');
		F_Note(bFailed := (rig.fbElev.bEnable OR rig.fbAzim.bEnable OR rig.fbDero.bEnable OR rig.fbBrakeHyd.BrakeOpen), sText := CONCAT(sTest, 'axes disabled, brake closed'));
		AssertFalse(Condition := bSawStop, Message := 'no stop at all');
		F_Note(bFailed := (bSawStop), sText := CONCAT(sTest, 'no stop at all'));
		AssertTrue(Condition := rig.fbTel.bCloseRoofRequest, Message := 'the roof request stays latched');
		F_Note(bFailed := NOT (rig.fbTel.bCloseRoofRequest), sText := CONCAT(sTest, 'the roof request stays latched'));
		rig.fbTel.Reset();
		nStep := 70;
		nCycles := 0;
	ELSIF nCycles > 600 THEN
		AssertTrue(Condition := FALSE, Message := 'the park after the release did not finish');
		F_Note(bFailed := TRUE, sText := CONCAT(sTest, 'the park after the release did not finish'));
		nStep := 99;
		TEST_FINISHED();
	END_IF
70:
	IF nCycles >= 10 THEN
		AssertFalse(Condition := rig.fbTel.bCloseRoofRequest, Message := 'the reset after the release clears the roof request');
		F_Note(bFailed := (rig.fbTel.bCloseRoofRequest), sText := CONCAT(sTest, 'the reset after the release clears the roof request'));
		rig.fbTel.Init();
		nStep := 80;
		nCycles := 0;
	END_IF
80:	// power=1: online again
	IF rig.Online THEN
		AssertTrue(Condition := TRUE, Message := 'online again after the release, the reset and power=1');
		nStep := 99;
		TEST_FINISHED();
	ELSIF nCycles > 1500 THEN
		AssertTrue(Condition := FALSE, Message := 'not online again after the release, the reset and power=1');
		F_Note(bFailed := TRUE, sText := CONCAT(sTest, 'not online again after the release, the reset and power=1'));
		nStep := 99;
		TEST_FINISHED();
	END_IF
END_CASE
END_METHOD

// #24 step 7 PR 6 (D8, row safety error; until 0.13.0 a safety error without E-stop only acted on the brake in the Wake&Shake window):
// a safety error (SafetyHandling.error, no E-stop) under tracking is handled as the E-stop: in its scan the axes are disabled and the
// hydraulics switched off (the lock is the stop, no bStop, no MC_Stop), tracking ends; nothing parks and the covers are not
// commanded while it is there (it is not bError); the roof close is requested. When it is gone the held park runs in place.
METHOD PRIVATE Safety_Error_While_Tracking_Locks_Then_Parks_In_Place_When_It_Clears
VAR_INST
	rig			: FB_MonetRig;
	nStep		: INT;
	nCycles		: UINT;
	nTracking	: UINT;
	sTest		: STRING(80);
	nDisable0	: UINT;	// hydraulics-off writes before the safety error
	nDisable1	: UINT;	// ... before it clears
	nEdges0		: UINT;	// MC_Stop requests of the three axes before the safety error
	bSawStop	: BOOL;
END_VAR
TEST('Safety_Error_While_Tracking_Locks_Then_Parks_In_Place_When_It_Clears');
sTest := 'Safety_Error_While_Tracking_Locks_Then_Parks_In_Place_When_It_Clears: ';
IF nStep >= 90 THEN
	RETURN;
END_IF
rig.Scan();
nCycles := nCycles + 1;
CASE nStep OF
0:	// wait for the clock, then power on
	IF rig.ClockValid THEN
		rig.fbTel.Init();
		nStep := 10;
		nCycles := 0;
	ELSIF nCycles > 2000 THEN
		AssertTrue(Condition := FALSE, Message := 'the astronomical clock never became valid');
		F_Note(bFailed := TRUE, sText := CONCAT(sTest, 'the astronomical clock never became valid'));
		nStep := 99;
		TEST_FINISHED();
	END_IF
10:	// online: track a circumpolar target
	IF rig.Online THEN
		rig.fbTel.Track(fRightAscension := 0.0, fDeclination := -85.0);
		nStep := 20;
		nCycles := 0;
	ELSIF nCycles > 1500 THEN
		AssertTrue(Condition := FALSE, Message := 'the mock telescope did not reach READY_STATE 1.0');
		F_Note(bFailed := TRUE, sText := CONCAT(sTest, 'the mock telescope did not reach READY_STATE 1.0'));
		nStep := 99;
		TEST_FINISHED();
	END_IF
20:	// tracking: the safety error comes
	IF rig.fbAzim.Tracking AND rig.fbElev.Tracking AND rig.fbDero.Tracking THEN
		nTracking := nTracking + 1;
	ELSE
		nTracking := 0;
	END_IF
	IF nTracking >= 5 THEN
		nDisable0 := rig.fbBrakeHyd.nDisableCalls;
		nEdges0 := rig.fbElev.nStopEdges + rig.fbAzim.nStopEdges + rig.fbDero.nStopEdges;
		rig.SetSafetyError(TRUE);
		nStep := 30;
		nCycles := 0;
	ELSIF nCycles > 800 THEN
		AssertTrue(Condition := FALSE, Message := 'the telescope did not start tracking');
		F_Note(bFailed := TRUE, sText := CONCAT(sTest, 'the telescope did not start tracking'));
		nStep := 99;
		TEST_FINISHED();
	END_IF
30:	// the lock is the stop; the park is held while the safety error is there
	bSawStop := bSawStop OR rig.fbTel.bStopActive;
	IF nCycles = 1 THEN	// the scan that saw the safety error
		AssertFalse(Condition := rig.fbElev.bEnable OR rig.fbAzim.bEnable OR rig.fbDero.bEnable, Message := 'the axes are disabled in the scan of the safety error');
		F_Note(bFailed := (rig.fbElev.bEnable OR rig.fbAzim.bEnable OR rig.fbDero.bEnable), sText := CONCAT(sTest, 'the axes are disabled in the scan of the safety error'));
		AssertTrue(Condition := rig.fbBrakeHyd.nDisableCalls > nDisable0, Message := 'the hydraulics go off in the scan of the safety error');
		F_Note(bFailed := NOT (rig.fbBrakeHyd.nDisableCalls > nDisable0), sText := CONCAT(sTest, 'the hydraulics go off in the scan of the safety error'));
		AssertTrue(Condition := rig.fbCovers.nStopCalls >= 1, Message := 'the covers get Stop() in the scan of the safety error (not on the E-stop circuit)');
		F_Note(bFailed := NOT (rig.fbCovers.nStopCalls >= 1), sText := CONCAT(sTest, 'the covers get Stop() in the scan of the safety error (not on the E-stop circuit)'));
	END_IF
	IF nCycles >= 30 THEN
		AssertFalse(Condition := rig.fbTel.bTrackActive OR rig.fbAzim.Tracking OR rig.fbElev.Tracking OR rig.fbDero.Tracking, Message := 'tracking has ended');
		F_Note(bFailed := (rig.fbTel.bTrackActive OR rig.fbAzim.Tracking OR rig.fbElev.Tracking OR rig.fbDero.Tracking), sText := CONCAT(sTest, 'tracking has ended'));
		AssertFalse(Condition := rig.fbElev.bEnable OR rig.fbAzim.bEnable OR rig.fbDero.bEnable, Message := 'the three axes stay disabled');
		F_Note(bFailed := (rig.fbElev.bEnable OR rig.fbAzim.bEnable OR rig.fbDero.bEnable), sText := CONCAT(sTest, 'the three axes stay disabled'));
		AssertFalse(Condition := rig.fbTel.bParkActive OR rig.fbTel.bIsParked, Message := 'no park while the safety error is there');
		F_Note(bFailed := (rig.fbTel.bParkActive OR rig.fbTel.bIsParked), sText := CONCAT(sTest, 'no park while the safety error is there'));
		AssertTrue(Condition := rig.fbCovers.nCloseCalls = 0, Message := 'the covers are not commanded while the safety error is there');
		F_Note(bFailed := NOT (rig.fbCovers.nCloseCalls = 0), sText := CONCAT(sTest, 'the covers are not commanded while the safety error is there'));
		AssertFalse(Condition := rig.fbTel.bError, Message := 'the safety error is not bError');
		F_Note(bFailed := (rig.fbTel.bError), sText := CONCAT(sTest, 'the safety error is not bError'));
		AssertTrue(Condition := rig.fbTel.bCloseRoofRequest, Message := 'the roof close is requested');
		F_Note(bFailed := NOT (rig.fbTel.bCloseRoofRequest), sText := CONCAT(sTest, 'the roof close is requested'));
		nDisable1 := rig.fbBrakeHyd.nDisableCalls;
		rig.SetSafetyError(FALSE);
		nStep := 40;
		nCycles := 0;
	END_IF
40:	// the safety error is gone: the park in place
	bSawStop := bSawStop OR rig.fbTel.bStopActive;
	IF rig.fbTel.bIsParked AND nCycles > 5 THEN
		AssertTrue(Condition := rig.fbTel.bParkedInPlace AND NOT rig.fbTel.bParkActive, Message := 'the park ended in place');
		F_Note(bFailed := NOT (rig.fbTel.bParkedInPlace AND NOT rig.fbTel.bParkActive), sText := CONCAT(sTest, 'the park ended in place'));
		AssertTrue(Condition := rig.fbCovers.bClosed AND rig.fbCovers.nCloseCalls >= 1, Message := 'the covers are closed');
		F_Note(bFailed := NOT (rig.fbCovers.bClosed AND rig.fbCovers.nCloseCalls >= 1), sText := CONCAT(sTest, 'the covers are closed'));
		AssertTrue(Condition := rig.fbBrakeHyd.nDisableCalls > nDisable1, Message := 'the park switches the hydraulics off');
		F_Note(bFailed := NOT (rig.fbBrakeHyd.nDisableCalls > nDisable1), sText := CONCAT(sTest, 'the park switches the hydraulics off'));
		AssertFalse(Condition := rig.fbBrakeHyd.BrakeOpen, Message := 'the brake is closed');
		F_Note(bFailed := (rig.fbBrakeHyd.BrakeOpen), sText := CONCAT(sTest, 'the brake is closed'));
		AssertFalse(Condition := bSawStop, Message := 'no ramp (bStop never set)');
		F_Note(bFailed := (bSawStop), sText := CONCAT(sTest, 'no ramp (bStop never set)'));
		AssertTrue(Condition := rig.fbElev.nStopEdges + rig.fbAzim.nStopEdges + rig.fbDero.nStopEdges = nEdges0, Message := 'no MC_Stop was sent');
		F_Note(bFailed := NOT (rig.fbElev.nStopEdges + rig.fbAzim.nStopEdges + rig.fbDero.nStopEdges = nEdges0), sText := CONCAT(sTest, 'no MC_Stop was sent'));
		nStep := 99;
		TEST_FINISHED();
	ELSIF nCycles > 600 THEN
		AssertTrue(Condition := FALSE, Message := 'the park did not finish after the safety error');
		F_Note(bFailed := TRUE, sText := CONCAT(sTest, 'the park did not finish after the safety error'));
		nStep := 99;
		TEST_FINISHED();
	END_IF
END_CASE
END_METHOD

// #24 step 7 PR 7 (D8, row power failure; until 0.13.0 Power_Failure_During_Goto_Keeps_Moving_Current: READY_STATE -2.0, the goto
// went on): bMainReady FALSE (MAIN: PowerMonitoring.phaseOK) during a goto is a telescope error (bHwError) and, with the drives still
// able to ramp on the mock (brake open, pressure there, no axis error), ramps first: in the scan of the failure bStop is set and the
// axes stay enabled; every axis is sent its MC_Stop while still enabled. After the stop has settled the queued emergency park parks in
// place: axes disabled, brake closed, covers closed, hydraulics off, bIsParked, bParkedInPlace; READY_STATE -1.0 and bCloseRoofRequest
// while the failure lasts. When the supply is back bError drops by itself, READY_STATE 0.0 (parked), not online without a new Init.
// What the drives do on a real phase loss is not modelled.
METHOD PRIVATE Power_Failure_During_Goto_Ramps_Then_Parks_In_Place
VAR_INST
	rig			: FB_MonetRig;
	nStep		: INT;
	nCycles		: UINT;
	sTest		: STRING(80);
	nEl0		: UINT;	// stop edges per axis before the failure
	nAz0		: UINT;
	nDr0		: UINT;
	nExt0		: UINT;	// 0x4257 rejections of the three axes before the failure
	nEdgesLast	: UINT;
	nEdgesNow	: UINT;
	nDisable0	: UINT;
	bSawStop	: BOOL;
	bStopOnDisabled	: BOOL;	// a stop edge came in a scan in which an axis was already disabled
END_VAR
TEST('Power_Failure_During_Goto_Ramps_Then_Parks_In_Place');
sTest := 'Power_Failure_During_Goto_Ramps_Then_Parks_In_Place: ';
IF nStep >= 90 THEN
	RETURN;
END_IF
rig.Scan();
nCycles := nCycles + 1;
CASE nStep OF
0:	// wait for the clock, then power on
	IF rig.ClockValid THEN
		rig.fbTel.Init();
		nStep := 10;
		nCycles := 0;
	ELSIF nCycles > 2000 THEN
		AssertTrue(Condition := FALSE, Message := 'the astronomical clock never became valid');
		F_Note(bFailed := TRUE, sText := CONCAT(sTest, 'the astronomical clock never became valid'));
		nStep := 99;
		TEST_FINISHED();
	END_IF
10:	// online: slow axes, goto a circumpolar target
	IF rig.Online THEN
		rig.SetMoveScans(nScans := 3000);
		rig.fbTel.Track(fRightAscension := 0.0, fDeclination := -85.0);
		nStep := 20;
		nCycles := 0;
	ELSIF nCycles > 1500 THEN
		AssertTrue(Condition := FALSE, Message := 'the mock telescope did not reach READY_STATE 1.0');
		F_Note(bFailed := TRUE, sText := CONCAT(sTest, 'the mock telescope did not reach READY_STATE 1.0'));
		nStep := 99;
		TEST_FINISHED();
	END_IF
20:
	IF rig.fbElev.MoveAxis AND rig.fbAzim.MoveAxis AND rig.fbDero.MoveAxis THEN
		nStep := 30;
		nCycles := 0;
	ELSIF nCycles > 300 THEN
		AssertTrue(Condition := FALSE, Message := 'the goto did not start the axis moves');
		F_Note(bFailed := TRUE, sText := CONCAT(sTest, 'the goto did not start the axis moves'));
		nStep := 99;
		TEST_FINISHED();
	END_IF
30:	// the axes move: the main power fails
	IF nCycles >= 5 THEN
		nEl0 := rig.fbElev.nStopEdges;
		nAz0 := rig.fbAzim.nStopEdges;
		nDr0 := rig.fbDero.nStopEdges;
		nEdgesLast := nEl0 + nAz0 + nDr0;
		nExt0 := rig.fbElev.nExtErrors + rig.fbAzim.nExtErrors + rig.fbDero.nExtErrors;
		nDisable0 := rig.fbBrakeHyd.nDisableCalls;
		rig.SetMainReady(FALSE);
		nStep := 40;
		nCycles := 0;
	END_IF
40:	// ramp, then the park in place
	bSawStop := bSawStop OR rig.fbTel.bStopActive;
	nEdgesNow := rig.fbElev.nStopEdges + rig.fbAzim.nStopEdges + rig.fbDero.nStopEdges;
	IF nEdgesNow > nEdgesLast AND NOT (rig.fbElev.bEnable AND rig.fbAzim.bEnable AND rig.fbDero.bEnable) THEN
		bStopOnDisabled := TRUE;
	END_IF
	nEdgesLast := nEdgesNow;
	IF nCycles = 1 THEN	// the scan that saw the failure
		AssertTrue(Condition := rig.fbTel.bStopActive AND rig.fbTel.bError, Message := 'the failure stops the axes in its scan (bStop) and is a telescope error');
		F_Note(bFailed := NOT (rig.fbTel.bStopActive AND rig.fbTel.bError), sText := CONCAT(sTest, 'the failure stops the axes in its scan (bStop) and is a telescope error'));
		AssertTrue(Condition := rig.fbElev.bEnable AND rig.fbAzim.bEnable AND rig.fbDero.bEnable, Message := 'the axes stay enabled for the ramp');
		F_Note(bFailed := NOT (rig.fbElev.bEnable AND rig.fbAzim.bEnable AND rig.fbDero.bEnable), sText := CONCAT(sTest, 'the axes stay enabled for the ramp'));
	END_IF
	IF rig.fbTel.bIsParked AND nCycles > 5 THEN
		AssertTrue(Condition := bSawStop, Message := 'the power failure ramped (bStop)');
		F_Note(bFailed := NOT (bSawStop), sText := CONCAT(sTest, 'the power failure ramped (bStop)'));
		AssertTrue(Condition := rig.fbElev.nStopEdges > nEl0 AND rig.fbAzim.nStopEdges > nAz0 AND rig.fbDero.nStopEdges > nDr0, Message := 'every axis was sent its MC_Stop');
		F_Note(bFailed := NOT (rig.fbElev.nStopEdges > nEl0 AND rig.fbAzim.nStopEdges > nAz0 AND rig.fbDero.nStopEdges > nDr0), sText := CONCAT(sTest, 'every axis was sent its MC_Stop'));
		AssertFalse(Condition := bStopOnDisabled, Message := 'the stops came before the disable');
		F_Note(bFailed := (bStopOnDisabled), sText := CONCAT(sTest, 'the stops came before the disable'));
		AssertTrue(Condition := rig.fbElev.nExtErrors + rig.fbAzim.nExtErrors + rig.fbDero.nExtErrors = nExt0, Message := 'no stop met the setpoint generator (0x4257)');
		F_Note(bFailed := NOT (rig.fbElev.nExtErrors + rig.fbAzim.nExtErrors + rig.fbDero.nExtErrors = nExt0), sText := CONCAT(sTest, 'no stop met the setpoint generator (0x4257)'));
		AssertTrue(Condition := rig.fbTel.bParkedInPlace AND NOT rig.fbTel.bParkActive, Message := 'the park ended in place');
		F_Note(bFailed := NOT (rig.fbTel.bParkedInPlace AND NOT rig.fbTel.bParkActive), sText := CONCAT(sTest, 'the park ended in place'));
		AssertFalse(Condition := rig.fbElev.bEnable OR rig.fbAzim.bEnable OR rig.fbDero.bEnable, Message := 'all three axes are disabled');
		F_Note(bFailed := (rig.fbElev.bEnable OR rig.fbAzim.bEnable OR rig.fbDero.bEnable), sText := CONCAT(sTest, 'all three axes are disabled'));
		AssertFalse(Condition := rig.fbBrakeHyd.BrakeOpen, Message := 'the brake is closed');
		F_Note(bFailed := (rig.fbBrakeHyd.BrakeOpen), sText := CONCAT(sTest, 'the brake is closed'));
		AssertTrue(Condition := rig.fbCovers.bClosed AND rig.fbCovers.nCloseCalls >= 1, Message := 'the covers are closed');
		F_Note(bFailed := NOT (rig.fbCovers.bClosed AND rig.fbCovers.nCloseCalls >= 1), sText := CONCAT(sTest, 'the covers are closed'));
		AssertTrue(Condition := rig.fbBrakeHyd.nDisableCalls > nDisable0, Message := 'the hydraulics are switched off');
		F_Note(bFailed := NOT (rig.fbBrakeHyd.nDisableCalls > nDisable0), sText := CONCAT(sTest, 'the hydraulics are switched off'));
		AssertFalse(Condition := rig.fbTel.bGotoActive OR rig.fbTel.bTrackActive, Message := 'the goto and the track are dropped');
		F_Note(bFailed := (rig.fbTel.bGotoActive OR rig.fbTel.bTrackActive), sText := CONCAT(sTest, 'the goto and the track are dropped'));
		AssertTrue(Condition := rig.fbTel.bError AND rig.fbTel.ReadyState = -1.0, Message := 'the failure is a telescope error, READY_STATE -1.0');
		F_Note(bFailed := NOT (rig.fbTel.bError AND rig.fbTel.ReadyState = -1.0), sText := CONCAT(sTest, 'the failure is a telescope error, READY_STATE -1.0'));
		AssertTrue(Condition := rig.fbTel.bCloseRoofRequest, Message := 'the roof close is requested');
		F_Note(bFailed := NOT (rig.fbTel.bCloseRoofRequest), sText := CONCAT(sTest, 'the roof close is requested'));
		rig.SetMainReady(TRUE);
		nStep := 50;
		nCycles := 0;
	ELSIF nCycles > 800 THEN
		AssertTrue(Condition := FALSE, Message := 'the telescope did not park after the ramp');
		F_Note(bFailed := TRUE, sText := CONCAT(sTest, 'the telescope did not park after the ramp'));
		nStep := 99;
		TEST_FINISHED();
	END_IF
50:	// the supply is back
	IF nCycles >= 10 THEN
		AssertFalse(Condition := rig.fbTel.bError, Message := 'bError drops by itself when the supply is back');
		F_Note(bFailed := (rig.fbTel.bError), sText := CONCAT(sTest, 'bError drops by itself when the supply is back'));
		AssertTrue(Condition := rig.fbTel.bIsParked AND rig.fbTel.ReadyState = 0.0 AND NOT rig.Online, Message := 'parked (READY_STATE 0.0), not online without a new Init');
		F_Note(bFailed := NOT (rig.fbTel.bIsParked AND rig.fbTel.ReadyState = 0.0 AND NOT rig.Online), sText := CONCAT(sTest, 'parked (READY_STATE 0.0), not online without a new Init'));
		nStep := 99;
		TEST_FINISHED();
	END_IF
END_CASE
END_METHOD

// #24 step 7 PR 7 (D8, row power failure): a phase loss that also stops the hydraulic pump (mock InjectPressureLoss in the same scan:
// the brake locks, the hydraulics report an error) leaves nothing that can ramp, the brake lock is the stop: the axes are disabled in
// the scan of the failure, bStop is never set, no MC_Stop is sent, and the emergency park parks in place (covers closed, hydraulics
// off, bIsParked, bParkedInPlace). Checks that the ramp of the power failure also asks whether the drives can still ramp.
METHOD PRIVATE Power_Failure_With_Pressure_Loss_Parks_In_Place_Without_Ramp
VAR_INST
	rig			: FB_MonetRig;
	nStep		: INT;
	nCycles		: UINT;
	nTracking	: UINT;
	sTest		: STRING(80);
	nEdges0		: UINT;	// stop edges of the three axes before the failure
	nDisable0	: UINT;
	bSawStop	: BOOL;
END_VAR
TEST('Power_Failure_With_Pressure_Loss_Parks_In_Place_Without_Ramp');
sTest := 'Power_Failure_With_Pressure_Loss_Parks_In_Place_Without_Ramp: ';
IF nStep >= 90 THEN
	RETURN;
END_IF
rig.Scan();
nCycles := nCycles + 1;
CASE nStep OF
0:	// wait for the clock, then power on
	IF rig.ClockValid THEN
		rig.fbTel.Init();
		nStep := 10;
		nCycles := 0;
	ELSIF nCycles > 2000 THEN
		AssertTrue(Condition := FALSE, Message := 'the astronomical clock never became valid');
		F_Note(bFailed := TRUE, sText := CONCAT(sTest, 'the astronomical clock never became valid'));
		nStep := 99;
		TEST_FINISHED();
	END_IF
10:	// online: track a circumpolar target
	IF rig.Online THEN
		rig.fbTel.Track(fRightAscension := 0.0, fDeclination := -85.0);
		nStep := 20;
		nCycles := 0;
	ELSIF nCycles > 1500 THEN
		AssertTrue(Condition := FALSE, Message := 'the mock telescope did not reach READY_STATE 1.0');
		F_Note(bFailed := TRUE, sText := CONCAT(sTest, 'the mock telescope did not reach READY_STATE 1.0'));
		nStep := 99;
		TEST_FINISHED();
	END_IF
20:	// tracking: the phase fails and with it the oil pressure (the brake locks)
	IF rig.fbAzim.Tracking AND rig.fbElev.Tracking AND rig.fbDero.Tracking THEN
		nTracking := nTracking + 1;
	ELSE
		nTracking := 0;
	END_IF
	IF nTracking >= 5 THEN
		nEdges0 := rig.fbElev.nStopEdges + rig.fbAzim.nStopEdges + rig.fbDero.nStopEdges;
		nDisable0 := rig.fbBrakeHyd.nDisableCalls;
		rig.SetMainReady(FALSE);
		rig.fbBrakeHyd.InjectPressureLoss();
		nStep := 30;
		nCycles := 0;
	ELSIF nCycles > 800 THEN
		AssertTrue(Condition := FALSE, Message := 'the telescope did not start tracking');
		F_Note(bFailed := TRUE, sText := CONCAT(sTest, 'the telescope did not start tracking'));
		nStep := 99;
		TEST_FINISHED();
	END_IF
30:
	bSawStop := bSawStop OR rig.fbTel.bStopActive;
	IF nCycles = 1 THEN	// the scan that saw the failure
		AssertFalse(Condition := rig.fbElev.bEnable OR rig.fbAzim.bEnable OR rig.fbDero.bEnable, Message := 'the lock is the stop: disabled in the scan of the failure');
		F_Note(bFailed := (rig.fbElev.bEnable OR rig.fbAzim.bEnable OR rig.fbDero.bEnable), sText := CONCAT(sTest, 'the lock is the stop: disabled in the scan of the failure'));
	END_IF
	IF rig.fbTel.bIsParked AND nCycles > 5 THEN
		AssertFalse(Condition := bSawStop, Message := 'no ramp (bStop never set)');
		F_Note(bFailed := (bSawStop), sText := CONCAT(sTest, 'no ramp (bStop never set)'));
		AssertTrue(Condition := rig.fbElev.nStopEdges + rig.fbAzim.nStopEdges + rig.fbDero.nStopEdges = nEdges0, Message := 'no MC_Stop was sent');
		F_Note(bFailed := NOT (rig.fbElev.nStopEdges + rig.fbAzim.nStopEdges + rig.fbDero.nStopEdges = nEdges0), sText := CONCAT(sTest, 'no MC_Stop was sent'));
		AssertTrue(Condition := rig.fbTel.bParkedInPlace AND NOT rig.fbTel.bParkActive, Message := 'the park ended in place');
		F_Note(bFailed := NOT (rig.fbTel.bParkedInPlace AND NOT rig.fbTel.bParkActive), sText := CONCAT(sTest, 'the park ended in place'));
		AssertTrue(Condition := rig.fbCovers.bClosed AND rig.fbBrakeHyd.nDisableCalls > nDisable0, Message := 'covers closed, hydraulics switched off');
		F_Note(bFailed := NOT (rig.fbCovers.bClosed AND rig.fbBrakeHyd.nDisableCalls > nDisable0), sText := CONCAT(sTest, 'covers closed, hydraulics switched off'));
		AssertTrue(Condition := rig.fbTel.bError AND rig.fbTel.ReadyState = -1.0 AND rig.fbTel.bCloseRoofRequest, Message := 'READY_STATE -1.0, roof close requested');
		F_Note(bFailed := NOT (rig.fbTel.bError AND rig.fbTel.ReadyState = -1.0 AND rig.fbTel.bCloseRoofRequest), sText := CONCAT(sTest, 'READY_STATE -1.0, roof close requested'));
		nStep := 99;
		TEST_FINISHED();
	ELSIF nCycles > 800 THEN
		AssertTrue(Condition := FALSE, Message := 'the emergency park did not finish');
		F_Note(bFailed := TRUE, sText := CONCAT(sTest, 'the emergency park did not finish'));
		nStep := 99;
		TEST_FINISHED();
	END_IF
END_CASE
END_METHOD

// #24 step 7 PR 5 (D8, row software error timeout; until 0.13.0 Goto_Times_Out_Without_Park_Current, which pinned the disable under
// motion without a park): a goto still running after 600 s is software error 16#10 (time seam: 1000, so 0.6 s). In the next scan the
// timeout ramps: bStop (stop transaction, #96) with the axes still enabled, one MC_Stop per axis before any disable. After the stop
// has settled the park queued behind it (bParkAfterStop) drives to the park position (el 60, az 175 of the rig), then disables the
// axes, closes the brake and the covers and switches the hydraulics off: bIsParked, not bParkedInPlace. The error stays latched
// (READY_STATE -1.0) and there is no roof close request (D9: recoverable).
METHOD PRIVATE Goto_Times_Out_Ramps_Then_Drives_To_Park
VAR_INST
	rig			: FB_MonetRig;
	nStep		: INT;
	nCycles		: UINT;
	sTest		: STRING(80);
	nEl0		: UINT;	// stop edges per axis before the ramp
	nAz0		: UINT;
	nDr0		: UINT;
	nEdgesLast	: UINT;
	nEdgesNow	: UINT;
	nDisable0	: UINT;
	nCoverClose0	: UINT;
	bSawStop	: BOOL;
	bStopOnDisabled	: BOOL;	// a stop edge came in a scan in which an axis was already disabled
	bParkMoveScans	: BOOL;	// the park move got the default 60 scans
END_VAR
TEST('Goto_Times_Out_Ramps_Then_Drives_To_Park');
sTest := 'Goto_Times_Out_Ramps_Then_Drives_To_Park: ';
IF nStep >= 90 THEN
	RETURN;
END_IF
rig.Scan();
nCycles := nCycles + 1;
CASE nStep OF
0:	// wait for the clock, then power on
	IF rig.ClockValid THEN
		rig.fbTel.Init();
		nStep := 10;
		nCycles := 0;
	ELSIF nCycles > 2000 THEN
		AssertTrue(Condition := FALSE, Message := 'the astronomical clock never became valid');
		F_Note(bFailed := TRUE, sText := CONCAT(sTest, 'the astronomical clock never became valid'));
		rig.SetTimeDivisor(nValue := 1);
		nStep := 99;
		TEST_FINISHED();
	END_IF
10:	// online: slow axes, short timeouts, goto a circumpolar target
	IF rig.Online THEN
		rig.SetMoveScans(nScans := 60000);
		rig.SetTimeDivisor(nValue := 1000);
		rig.fbTel.Track(fRightAscension := 0.0, fDeclination := -85.0);
		nStep := 20;
		nCycles := 0;
	ELSIF nCycles > 1500 THEN
		AssertTrue(Condition := FALSE, Message := 'the mock telescope did not reach READY_STATE 1.0');
		F_Note(bFailed := TRUE, sText := CONCAT(sTest, 'the mock telescope did not reach READY_STATE 1.0'));
		rig.SetTimeDivisor(nValue := 1);
		nStep := 99;
		TEST_FINISHED();
	END_IF
20:
	IF rig.fbTel.bError THEN
		rig.SetTimeDivisor(nValue := 1);
		AssertTrue(Condition := rig.fbTel.nErrorID = 16#10, Message := 'the goto timeout is error 16#10');
		F_Note(bFailed := NOT (rig.fbTel.nErrorID = 16#10), sText := CONCAT(sTest, 'the goto timeout is error 16#10'));
		AssertFalse(Condition := rig.fbTel.bGotoActive, Message := 'the goto is dropped');
		F_Note(bFailed := (rig.fbTel.bGotoActive), sText := CONCAT(sTest, 'the goto is dropped'));
		nEl0 := rig.fbElev.nStopEdges;
		nAz0 := rig.fbAzim.nStopEdges;
		nDr0 := rig.fbDero.nStopEdges;
		nEdgesLast := nEl0 + nAz0 + nDr0;
		nDisable0 := rig.fbBrakeHyd.nDisableCalls;
		nCoverClose0 := rig.fbCovers.nCloseCalls;
		nStep := 30;
		nCycles := 0;
	ELSIF nCycles > 3000 THEN
		AssertTrue(Condition := FALSE, Message := 'the goto never timed out');
		F_Note(bFailed := TRUE, sText := CONCAT(sTest, 'the goto never timed out'));
		rig.SetTimeDivisor(nValue := 1);
		nStep := 99;
		TEST_FINISHED();
	END_IF
30:	// the ramp, then the park to the park position
	bSawStop := bSawStop OR rig.fbTel.bStopActive;
	nEdgesNow := rig.fbElev.nStopEdges + rig.fbAzim.nStopEdges + rig.fbDero.nStopEdges;
	IF nEdgesNow > nEdgesLast AND NOT (rig.fbElev.bEnable AND rig.fbAzim.bEnable AND rig.fbDero.bEnable) THEN
		bStopOnDisabled := TRUE;
	END_IF
	nEdgesLast := nEdgesNow;
	IF rig.fbTel.bParkActive AND NOT bParkMoveScans THEN	// the stop has settled (the goto move is aborted): the park move is a normal one
		rig.SetMoveScans(nScans := 60);
		bParkMoveScans := TRUE;
	END_IF
	IF nCycles = 1 THEN	// the scan after the one that raised the timeout
		AssertTrue(Condition := rig.fbTel.bStopActive AND rig.fbTel.bError, Message := 'the timeout stops the axes in the next scan (bStop)');
		F_Note(bFailed := NOT (rig.fbTel.bStopActive AND rig.fbTel.bError), sText := CONCAT(sTest, 'the timeout stops the axes in the next scan (bStop)'));
		AssertTrue(Condition := rig.fbElev.bEnable AND rig.fbAzim.bEnable AND rig.fbDero.bEnable, Message := 'the axes stay enabled for the ramp');
		F_Note(bFailed := NOT (rig.fbElev.bEnable AND rig.fbAzim.bEnable AND rig.fbDero.bEnable), sText := CONCAT(sTest, 'the axes stay enabled for the ramp'));
	END_IF
	IF rig.fbTel.bIsParked AND nCycles > 5 THEN
		AssertTrue(Condition := bSawStop AND rig.fbElev.nStopEdges > nEl0 AND rig.fbAzim.nStopEdges > nAz0 AND rig.fbDero.nStopEdges > nDr0, Message := 'the timeout ramped: every axis was sent its MC_Stop');
		F_Note(bFailed := NOT (bSawStop AND rig.fbElev.nStopEdges > nEl0 AND rig.fbAzim.nStopEdges > nAz0 AND rig.fbDero.nStopEdges > nDr0), sText := CONCAT(sTest, 'the timeout ramped: every axis was sent its MC_Stop'));
		AssertFalse(Condition := bStopOnDisabled, Message := 'the stops came before the disable');
		F_Note(bFailed := (bStopOnDisabled), sText := CONCAT(sTest, 'the stops came before the disable'));
		AssertTrue(Condition := NOT rig.fbTel.bParkedInPlace AND NOT rig.fbTel.bParkActive, Message := 'the park drove to the park position (not in place)');
		F_Note(bFailed := NOT (NOT rig.fbTel.bParkedInPlace AND NOT rig.fbTel.bParkActive), sText := CONCAT(sTest, 'the park drove to the park position (not in place)'));
		AssertTrue(Condition := ABS(rig.fbElev.fActualPosition - 60.0) < 0.001 AND ABS(rig.fbAzim.fActualPosition - 175.0) < 0.001, Message := 'the axes stand at the park position');
		F_Note(bFailed := NOT (ABS(rig.fbElev.fActualPosition - 60.0) < 0.001 AND ABS(rig.fbAzim.fActualPosition - 175.0) < 0.001), sText := CONCAT(sTest, 'the axes stand at the park position'));
		AssertFalse(Condition := rig.fbElev.bEnable OR rig.fbAzim.bEnable OR rig.fbDero.bEnable, Message := 'the three axes are disabled');
		F_Note(bFailed := (rig.fbElev.bEnable OR rig.fbAzim.bEnable OR rig.fbDero.bEnable), sText := CONCAT(sTest, 'the three axes are disabled'));
		AssertFalse(Condition := rig.fbBrakeHyd.BrakeOpen, Message := 'the brake is closed');
		F_Note(bFailed := (rig.fbBrakeHyd.BrakeOpen), sText := CONCAT(sTest, 'the brake is closed'));
		AssertTrue(Condition := rig.fbCovers.bClosed AND rig.fbCovers.nCloseCalls > nCoverClose0, Message := 'the covers are closed');
		F_Note(bFailed := NOT (rig.fbCovers.bClosed AND rig.fbCovers.nCloseCalls > nCoverClose0), sText := CONCAT(sTest, 'the covers are closed'));
		AssertTrue(Condition := rig.fbBrakeHyd.nDisableCalls > nDisable0, Message := 'the hydraulics are switched off');
		F_Note(bFailed := NOT (rig.fbBrakeHyd.nDisableCalls > nDisable0), sText := CONCAT(sTest, 'the hydraulics are switched off'));
		AssertTrue(Condition := rig.fbTel.bError AND rig.fbTel.nErrorID = 16#10 AND rig.fbTel.ReadyState = -1.0, Message := 'the error 16#10 is latched, READY_STATE -1.0');
		F_Note(bFailed := NOT (rig.fbTel.bError AND rig.fbTel.nErrorID = 16#10 AND rig.fbTel.ReadyState = -1.0), sText := CONCAT(sTest, 'the error 16#10 is latched, READY_STATE -1.0'));
		// step 7 PR 1 (D9): a software error is recoverable, no roof close request
		AssertFalse(Condition := rig.fbTel.bCloseRoofRequest, Message := 'no roof close request for 16#10');
		F_Note(bFailed := (rig.fbTel.bCloseRoofRequest), sText := CONCAT(sTest, 'no roof close request for 16#10'));
		nStep := 99;
		TEST_FINISHED();
	ELSIF nCycles > 1500 THEN
		AssertTrue(Condition := FALSE, Message := 'the telescope did not park after the timeout');
		F_Note(bFailed := TRUE, sText := CONCAT(sTest, 'the telescope did not park after the timeout'));
		nStep := 99;
		TEST_FINISHED();
	END_IF
END_CASE
END_METHOD

// #24 step 7 PR 5 (D8, row software error timeout; until 0.13.0 Home_Times_Out_Without_Park_Current): a home still running after
// 600 s is software error 16#30 (time seam: 1000, so 0.6 s); bGoHome is dropped. The same reaction as the goto timeout: in the next
// scan bStop with the axes enabled, then the park drives to the park position (el 60; the home position is el 40), axes disabled,
// brake and covers closed, hydraulics off, bIsParked, not bParkedInPlace; the error stays, no roof close request (D9).
METHOD PRIVATE Home_Times_Out_Ramps_Then_Drives_To_Park
VAR_INST
	rig			: FB_MonetRig;
	nStep		: INT;
	nCycles		: UINT;
	sTest		: STRING(80);
	nEdges0		: UINT;	// stop edges of the three axes before the ramp
	nDisable0	: UINT;
	nCoverClose0	: UINT;
	bSawStop	: BOOL;
	bParkMoveScans	: BOOL;	// the park move got the default 60 scans
END_VAR
TEST('Home_Times_Out_Ramps_Then_Drives_To_Park');
sTest := 'Home_Times_Out_Ramps_Then_Drives_To_Park: ';
IF nStep >= 90 THEN
	RETURN;
END_IF
rig.Scan();
nCycles := nCycles + 1;
CASE nStep OF
0:	// wait for the clock, then power on
	IF rig.ClockValid THEN
		rig.fbTel.Init();
		nStep := 10;
		nCycles := 0;
	ELSIF nCycles > 2000 THEN
		AssertTrue(Condition := FALSE, Message := 'the astronomical clock never became valid');
		F_Note(bFailed := TRUE, sText := CONCAT(sTest, 'the astronomical clock never became valid'));
		rig.SetTimeDivisor(nValue := 1);
		nStep := 99;
		TEST_FINISHED();
	END_IF
10:	// online: slow axes, short timeouts, home
	IF rig.Online THEN
		rig.SetMoveScans(nScans := 60000);
		rig.SetTimeDivisor(nValue := 1000);
		rig.fbTel.Home();
		nStep := 20;
		nCycles := 0;
	ELSIF nCycles > 1500 THEN
		AssertTrue(Condition := FALSE, Message := 'the mock telescope did not reach READY_STATE 1.0');
		F_Note(bFailed := TRUE, sText := CONCAT(sTest, 'the mock telescope did not reach READY_STATE 1.0'));
		rig.SetTimeDivisor(nValue := 1);
		nStep := 99;
		TEST_FINISHED();
	END_IF
20:
	IF rig.fbTel.bError THEN
		rig.SetTimeDivisor(nValue := 1);
		AssertTrue(Condition := rig.fbTel.nErrorID = 16#30, Message := 'the home timeout is error 16#30');
		F_Note(bFailed := NOT (rig.fbTel.nErrorID = 16#30), sText := CONCAT(sTest, 'the home timeout is error 16#30'));
		AssertFalse(Condition := rig.fbTel.bGoHomeActive, Message := 'the home is dropped');
		F_Note(bFailed := (rig.fbTel.bGoHomeActive), sText := CONCAT(sTest, 'the home is dropped'));
		nEdges0 := rig.fbElev.nStopEdges + rig.fbAzim.nStopEdges + rig.fbDero.nStopEdges;
		nDisable0 := rig.fbBrakeHyd.nDisableCalls;
		nCoverClose0 := rig.fbCovers.nCloseCalls;
		nStep := 30;
		nCycles := 0;
	ELSIF nCycles > 3000 THEN
		AssertTrue(Condition := FALSE, Message := 'the home never timed out');
		F_Note(bFailed := TRUE, sText := CONCAT(sTest, 'the home never timed out'));
		rig.SetTimeDivisor(nValue := 1);
		nStep := 99;
		TEST_FINISHED();
	END_IF
30:	// the ramp, then the park to the park position
	bSawStop := bSawStop OR rig.fbTel.bStopActive;
	IF rig.fbTel.bParkActive AND NOT bParkMoveScans THEN	// the stop has settled (the home move is aborted): the park move is a normal one
		rig.SetMoveScans(nScans := 60);
		bParkMoveScans := TRUE;
	END_IF
	IF nCycles = 1 THEN	// the scan after the one that raised the timeout
		AssertTrue(Condition := rig.fbTel.bStopActive AND rig.fbElev.bEnable AND rig.fbAzim.bEnable AND rig.fbDero.bEnable, Message := 'the timeout ramps (bStop) with the axes enabled');
		F_Note(bFailed := NOT (rig.fbTel.bStopActive AND rig.fbElev.bEnable AND rig.fbAzim.bEnable AND rig.fbDero.bEnable), sText := CONCAT(sTest, 'the timeout ramps (bStop) with the axes enabled'));
	END_IF
	IF rig.fbTel.bIsParked AND nCycles > 5 THEN
		AssertTrue(Condition := bSawStop AND rig.fbElev.nStopEdges + rig.fbAzim.nStopEdges + rig.fbDero.nStopEdges > nEdges0, Message := 'the timeout ramped (MC_Stop sent)');
		F_Note(bFailed := NOT (bSawStop AND rig.fbElev.nStopEdges + rig.fbAzim.nStopEdges + rig.fbDero.nStopEdges > nEdges0), sText := CONCAT(sTest, 'the timeout ramped (MC_Stop sent)'));
		AssertTrue(Condition := NOT rig.fbTel.bParkedInPlace AND ABS(rig.fbElev.fActualPosition - 60.0) < 0.001, Message := 'the park drove to the park position (el 60, not in place)');
		F_Note(bFailed := NOT (NOT rig.fbTel.bParkedInPlace AND ABS(rig.fbElev.fActualPosition - 60.0) < 0.001), sText := CONCAT(sTest, 'the park drove to the park position (el 60, not in place)'));
		AssertFalse(Condition := rig.fbElev.bEnable OR rig.fbAzim.bEnable OR rig.fbDero.bEnable, Message := 'the three axes are disabled');
		F_Note(bFailed := (rig.fbElev.bEnable OR rig.fbAzim.bEnable OR rig.fbDero.bEnable), sText := CONCAT(sTest, 'the three axes are disabled'));
		AssertFalse(Condition := rig.fbBrakeHyd.BrakeOpen, Message := 'the brake is closed');
		F_Note(bFailed := (rig.fbBrakeHyd.BrakeOpen), sText := CONCAT(sTest, 'the brake is closed'));
		AssertTrue(Condition := rig.fbCovers.bClosed AND rig.fbCovers.nCloseCalls > nCoverClose0, Message := 'the covers are closed');
		F_Note(bFailed := NOT (rig.fbCovers.bClosed AND rig.fbCovers.nCloseCalls > nCoverClose0), sText := CONCAT(sTest, 'the covers are closed'));
		AssertTrue(Condition := rig.fbBrakeHyd.nDisableCalls > nDisable0, Message := 'the hydraulics are switched off');
		F_Note(bFailed := NOT (rig.fbBrakeHyd.nDisableCalls > nDisable0), sText := CONCAT(sTest, 'the hydraulics are switched off'));
		AssertTrue(Condition := rig.fbTel.bError AND rig.fbTel.nErrorID = 16#30 AND rig.fbTel.ReadyState = -1.0, Message := 'the error 16#30 is latched, READY_STATE -1.0');
		F_Note(bFailed := NOT (rig.fbTel.bError AND rig.fbTel.nErrorID = 16#30 AND rig.fbTel.ReadyState = -1.0), sText := CONCAT(sTest, 'the error 16#30 is latched, READY_STATE -1.0'));
		AssertFalse(Condition := rig.fbTel.bCloseRoofRequest, Message := 'no roof close request for 16#30');
		F_Note(bFailed := (rig.fbTel.bCloseRoofRequest), sText := CONCAT(sTest, 'no roof close request for 16#30'));
		nStep := 99;
		TEST_FINISHED();
	ELSIF nCycles > 1500 THEN
		AssertTrue(Condition := FALSE, Message := 'the telescope did not park after the timeout');
		F_Note(bFailed := TRUE, sText := CONCAT(sTest, 'the telescope did not park after the timeout'));
		nStep := 99;
		TEST_FINISHED();
	END_IF
END_CASE
END_METHOD

// #24 step 5: the rising edge of the slew input while the clock is not valid is rejected with clock_invalid by the input gate
// (_CommandState, F_CommandAcceptance), like the Slew() method: no request is set, so the clock check of the body (a request while the
// clock is not valid sets bStopActive, the normal stop path) has nothing to stop and nothing parks. Until 0.14.x the written flag was
// seen by that check before the gate and also took the stop path (this test was Clock_Invalid_Slew_Takes_The_Stop_Path, same Id).
// Only reachable before the first clock sync: FB_AstroClockSync latches bValid. The input is written directly (an ADS write).
METHOD PRIVATE Clock_Invalid_Slew_Input_Is_Rejected
VAR_INST
	rig			: FB_MonetRig;
	nStep		: INT;
	nCycles		: UINT;
	sTest		: STRING(80);
	bSawStop	: BOOL;
END_VAR
TEST('Clock_Invalid_Slew_Input_Is_Rejected');
sTest := 'Clock_Invalid_Slew_Input_Is_Rejected: ';
IF nStep >= 90 THEN
	RETURN;
END_IF
rig.Scan();
nCycles := nCycles + 1;
CASE nStep OF
0:	// first cycle: the clock needs a NT_GetTime round trip (about 5 s), so it is not valid yet
	IF NOT rig.ClockValid THEN
		rig.SetSlewFlag();
		nStep := 10;
		nCycles := 0;
	ELSE
		AssertTrue(Condition := FALSE, Message := 'the clock was already valid in the first cycle');
		F_Note(bFailed := TRUE, sText := CONCAT(sTest, 'the clock was already valid in the first cycle'));
		nStep := 99;
		TEST_FINISHED();
	END_IF
10:
	bSawStop := bSawStop OR rig.fbTel.bStopActive;
	IF nCycles >= 10 THEN
		AssertFalse(Condition := rig.ClockValid, Message := 'the clock is still not valid');
		F_Note(bFailed := (rig.ClockValid), sText := CONCAT(sTest, 'the clock is still not valid'));
		AssertFalse(Condition := bSawStop, Message := 'the rejected slew input sets no request, so no stop');
		F_Note(bFailed := (bSawStop), sText := CONCAT(sTest, 'the rejected slew input sets no request, so no stop'));
		AssertFalse(Condition := rig.fbTel.bSlewActive, Message := 'the slew is dropped');
		F_Note(bFailed := (rig.fbTel.bSlewActive), sText := CONCAT(sTest, 'the slew is dropped'));
		AssertTrue(Condition := rig.fbTel.eLastRejectReason = MONETcommon.E_CommandRejectReason.clock_invalid, Message := 'the slew is rejected with clock_invalid');
		F_Note(bFailed := NOT (rig.fbTel.eLastRejectReason = MONETcommon.E_CommandRejectReason.clock_invalid), sText := CONCAT(sTest, 'the slew is rejected with clock_invalid'));
		AssertFalse(Condition := rig.fbTel.bParkActive OR rig.fbTel.bError, Message := 'no park, no error');
		F_Note(bFailed := (rig.fbTel.bParkActive OR rig.fbTel.bError), sText := CONCAT(sTest, 'no park, no error'));
		nStep := 99;
		TEST_FINISHED();
	END_IF
END_CASE
END_METHOD

// FB_MonetMqttWatchdog:29-35 (D4): armed only after the first connect; tGrace after the connection is lost it calls Park() on the
// telescope and Close() on the roof in the same scan, and again in every scan until the connection is back. The telescope is the
// real FB_MonetTelescopeControl of a rig whose body is not scanned here, so bPark stays as Park() set it; the roof is FB_RoofMock.
METHOD PRIVATE Watchdog_Parks_And_Closes_The_Roof_In_One_Scan
VAR_INST
	rig			: FB_MonetRig;
	fbRoof		: FB_RoofMock;
	bConnected	: BOOL;
	nStep		: INT;
	nCycles		: UINT;
	sTest		: STRING(80);
	nCloses		: UINT;
END_VAR
TEST('Watchdog_Parks_And_Closes_The_Roof_In_One_Scan');
sTest := 'Watchdog_Parks_And_Closes_The_Roof_In_One_Scan: ';
IF nStep >= 90 THEN
	RETURN;
END_IF
rig.fbWatchdog(bConnected := bConnected, iTelescope := rig.fbTel, iRoof := fbRoof, tGrace := T#100MS);
nCycles := nCycles + 1;
CASE nStep OF
0:	// never connected: not armed, also after more than tGrace; then the broker connects
	IF nCycles >= 30 THEN
		AssertFalse(Condition := rig.fbWatchdog.bTriggered OR rig.fbTel.bParkActive OR fbRoof.nCloseCalls > 0, Message := 'not armed before the first connect');
		F_Note(bFailed := (rig.fbWatchdog.bTriggered OR rig.fbTel.bParkActive OR fbRoof.nCloseCalls > 0), sText := CONCAT(sTest, 'not armed before the first connect'));
		bConnected := TRUE;
		nStep := 10;
		nCycles := 0;
	END_IF
10:	// connected for one scan, then the connection is lost
	bConnected := FALSE;
	nStep := 20;
	nCycles := 0;
20:
	IF rig.fbWatchdog.bTriggered THEN
		AssertTrue(Condition := rig.fbTel.bParkActive AND fbRoof.nCloseCalls = 1, Message := 'park and roof close in the trigger scan');
		F_Note(bFailed := NOT (rig.fbTel.bParkActive AND fbRoof.nCloseCalls = 1), sText := CONCAT(sTest, 'park and roof close in the trigger scan'));
		nStep := 30;
		nCycles := 0;
	ELSIF rig.fbTel.bParkActive OR fbRoof.nCloseCalls > 0 THEN
		AssertTrue(Condition := FALSE, Message := 'park or roof close before the watchdog triggered');
		F_Note(bFailed := TRUE, sText := CONCAT(sTest, 'park or roof close before the watchdog triggered'));
		nStep := 99;
		TEST_FINISHED();
	ELSIF nCycles > 300 THEN
		AssertTrue(Condition := FALSE, Message := 'the watchdog never triggered');
		F_Note(bFailed := TRUE, sText := CONCAT(sTest, 'the watchdog never triggered'));
		nStep := 99;
		TEST_FINISHED();
	END_IF
30:	// still disconnected: repeated in every scan; then the broker is back
	AssertTrue(Condition := fbRoof.nCloseCalls = 2, Message := 'the roof close is repeated in the next scan');
	F_Note(bFailed := NOT (fbRoof.nCloseCalls = 2), sText := CONCAT(sTest, 'the roof close is repeated in the next scan'));
	bConnected := TRUE;
	nStep := 40;
	nCycles := 0;
40:	// connected again: the watchdog lets go
	AssertFalse(Condition := rig.fbWatchdog.bTriggered, Message := 'not triggered once the connection is back');
	F_Note(bFailed := (rig.fbWatchdog.bTriggered), sText := CONCAT(sTest, 'not triggered once the connection is back'));
	nCloses := fbRoof.nCloseCalls;
	nStep := 50;
	nCycles := 0;
50:
	IF nCycles >= 10 THEN
		AssertTrue(Condition := fbRoof.nCloseCalls = nCloses, Message := 'no roof close while connected');
		F_Note(bFailed := NOT (fbRoof.nCloseCalls = nCloses), sText := CONCAT(sTest, 'no roof close while connected'));
		nStep := 99;
		TEST_FINISHED();
	END_IF
END_CASE
END_METHOD

// #24 step 2c, row "software error: config": an invalid stMotion (BROTLib.F_MotionConfigValid FALSE, here the goto window reversed,
// min 50 > max 40) is software error 16#32, raised in every scan like 16#31 (M: after F_HomeBelowHorizon). The defaults stay in use
// (stMotionUsed), a reset does not clear the error while the configuration is wrong, and it clears once the configuration is valid.
// No clock and no power-on needed.
METHOD PRIVATE Invalid_Motion_Config_Is_Software_Error_32
VAR_INST
	rig			: FB_MonetRig;
	stCfg		: BROTLib.ST_MotionConfig;
	stValid		: BROTLib.ST_MotionConfig;	// the defaults
	nStep		: INT;
	nCycles		: UINT;
	sTest		: STRING(80);
END_VAR
TEST('Invalid_Motion_Config_Is_Software_Error_32');
sTest := 'Invalid_Motion_Config_Is_Software_Error_32: ';
IF nStep >= 90 THEN
	RETURN;
END_IF
IF nStep = 0 THEN	// before the first scan
	stCfg.fGotoMinElevation := 50.0;
	stCfg.fGotoMaxElevation := 40.0;
	rig.SetMotion(stValue := stCfg);
	nStep := 10;
END_IF
rig.Scan();
nCycles := nCycles + 1;
CASE nStep OF
10:
	IF nCycles >= 3 THEN
		AssertTrue(Condition := rig.fbTel.bError AND rig.fbTel.nErrorID = 16#32, Message := 'the invalid configuration is error 16#32');
		F_Note(bFailed := NOT (rig.fbTel.bError AND rig.fbTel.nErrorID = 16#32), sText := CONCAT(sTest, 'the invalid configuration is error 16#32'));
		AssertTrue(Condition := rig.fbTel.stMotionUsed.fGotoMinElevation = 2.0 AND rig.fbTel.stMotionUsed.fGotoMaxElevation = 89.5,
			Message := 'the defaults stay in use');
		F_Note(bFailed := NOT (rig.fbTel.stMotionUsed.fGotoMinElevation = 2.0 AND rig.fbTel.stMotionUsed.fGotoMaxElevation = 89.5),
			sText := CONCAT(sTest, 'the defaults stay in use'));
		// step 7 PR 1 (D9): a configuration error is recoverable, no roof close request
		AssertFalse(Condition := rig.fbTel.bCloseRoofRequest, Message := 'no roof close request for 16#32');
		F_Note(bFailed := (rig.fbTel.bCloseRoofRequest), sText := CONCAT(sTest, 'no roof close request for 16#32'));
		rig.fbTel.Reset();
		nStep := 20;
		nCycles := 0;
	END_IF
20:
	IF nCycles >= 3 THEN
		AssertTrue(Condition := rig.fbTel.bError AND rig.fbTel.nErrorID = 16#32, Message := 'a reset does not clear it while the configuration is wrong');
		F_Note(bFailed := NOT (rig.fbTel.bError AND rig.fbTel.nErrorID = 16#32), sText := CONCAT(sTest, 'a reset does not clear it while the configuration is wrong'));
		rig.SetMotion(stValue := stValid);
		rig.fbTel.Reset();
		nStep := 30;
		nCycles := 0;
	END_IF
30:
	IF nCycles >= 3 THEN
		AssertFalse(Condition := rig.fbTel.bError, Message := 'a valid configuration and a reset clear the error');
		F_Note(bFailed := (rig.fbTel.bError), sText := CONCAT(sTest, 'a valid configuration and a reset clear the error'));
		nStep := 99;
		TEST_FINISHED();
	END_IF
END_CASE
END_METHOD

// #24 step 7 PR 1 (D9, row axis error): an elevation, azimuth and derotator error each set bCloseRoofRequest (M: next to bError).
// The axis error goes only with a reset: the telescope resets the axis in the reset scan (the cause is still active, the
// request stays), bReset is held while bError, so in the next scan the request is cleared without a second reset.
// No clock, no power-on (the telescope is parked at the start, so no emergency park).
METHOD PRIVATE Roof_Request_On_Axis_Errors
VAR_INST
	rig			: FB_MonetRig;
	nStep		: INT;
	nCycles		: UINT;
	sTest		: STRING(80);
END_VAR
TEST('Roof_Request_On_Axis_Errors');
sTest := 'Roof_Request_On_Axis_Errors: ';
IF nStep >= 90 THEN
	RETURN;
END_IF
rig.Scan();
nCycles := nCycles + 1;
// one step every 3 scans: the cause or the reset of the step before has been scanned
IF nCycles >= 3 THEN
	nCycles := 0;
	CASE nStep OF
	0:
		AssertFalse(Condition := rig.fbTel.bCloseRoofRequest, Message := 'no request without a cause');
		F_Note(bFailed := (rig.fbTel.bCloseRoofRequest), sText := CONCAT(sTest, 'no request without a cause'));
		rig.InjectElevationError(16#4550);
		nStep := 10;
	10:
		AssertTrue(Condition := rig.fbTel.bCloseRoofRequest, Message := 'the elevation error sets the request');
		F_Note(bFailed := NOT (rig.fbTel.bCloseRoofRequest), sText := CONCAT(sTest, 'the elevation error sets the request'));
		rig.fbTel.Reset();
		nStep := 20;
	20:
		AssertTrue(Condition := NOT rig.fbTel.bCloseRoofRequest AND NOT rig.fbTel.bError, Message := 'one reset clears the elevation error and the request');
		F_Note(bFailed := NOT (NOT rig.fbTel.bCloseRoofRequest AND NOT rig.fbTel.bError), sText := CONCAT(sTest, 'one reset clears the elevation error and the request'));
		rig.InjectAzimuthError(16#4550);
		nStep := 30;
	30:
		AssertTrue(Condition := rig.fbTel.bCloseRoofRequest, Message := 'the azimuth error sets the request');
		F_Note(bFailed := NOT (rig.fbTel.bCloseRoofRequest), sText := CONCAT(sTest, 'the azimuth error sets the request'));
		rig.fbTel.Reset();
		nStep := 40;
	40:
		AssertTrue(Condition := NOT rig.fbTel.bCloseRoofRequest AND NOT rig.fbTel.bError, Message := 'one reset clears the azimuth error and the request');
		F_Note(bFailed := NOT (NOT rig.fbTel.bCloseRoofRequest AND NOT rig.fbTel.bError), sText := CONCAT(sTest, 'one reset clears the azimuth error and the request'));
		rig.InjectDerotatorError(16#4550);
		nStep := 50;
	50:
		AssertTrue(Condition := rig.fbTel.bCloseRoofRequest, Message := 'the derotator error sets the request');
		F_Note(bFailed := NOT (rig.fbTel.bCloseRoofRequest), sText := CONCAT(sTest, 'the derotator error sets the request'));
		rig.fbTel.Reset();
		nStep := 60;
	60:
		AssertTrue(Condition := NOT rig.fbTel.bCloseRoofRequest AND NOT rig.fbTel.bError, Message := 'one reset clears the derotator error and the request');
		F_Note(bFailed := NOT (NOT rig.fbTel.bCloseRoofRequest AND NOT rig.fbTel.bError), sText := CONCAT(sTest, 'one reset clears the derotator error and the request'));
		nStep := 99;
		TEST_FINISHED();
	END_CASE
END_IF
END_METHOD

// #24 step 7 PR 1 (D9, row hydraulics error): fbHydraulics.Error sets bCloseRoofRequest although it is no telescope error. The
// telescope reset does not reset the hydraulics (HalfBROT Reset(), the MAIN reset button), so a reset with the error still
// there keeps the request; after the hydraulics reset it stays latched until the next telescope reset.
METHOD PRIVATE Roof_Request_On_Hydraulics_Error
VAR_INST
	rig			: FB_MonetRig;
	nStep		: INT;
	nCycles		: UINT;
	sTest		: STRING(80);
END_VAR
TEST('Roof_Request_On_Hydraulics_Error');
sTest := 'Roof_Request_On_Hydraulics_Error: ';
IF nStep >= 90 THEN
	RETURN;
END_IF
rig.Scan();
nCycles := nCycles + 1;
// one step every 3 scans: the cause or the reset of the step before has been scanned
IF nCycles >= 3 THEN
	nCycles := 0;
	CASE nStep OF
	0:
		AssertFalse(Condition := rig.fbTel.bCloseRoofRequest, Message := 'no request without a cause');
		F_Note(bFailed := (rig.fbTel.bCloseRoofRequest), sText := CONCAT(sTest, 'no request without a cause'));
		rig.fbBrakeHyd.InjectError();
		nStep := 10;
	10:
		AssertTrue(Condition := rig.fbTel.bCloseRoofRequest, Message := 'the hydraulics error sets the request');
		F_Note(bFailed := NOT (rig.fbTel.bCloseRoofRequest), sText := CONCAT(sTest, 'the hydraulics error sets the request'));
		rig.fbTel.Reset();
		nStep := 20;
	20:
		AssertTrue(Condition := rig.fbTel.bCloseRoofRequest, Message := 'a reset with the hydraulics error keeps it');
		F_Note(bFailed := NOT (rig.fbTel.bCloseRoofRequest), sText := CONCAT(sTest, 'a reset with the hydraulics error keeps it'));
		rig.fbBrakeHyd.Reset();
		nStep := 30;
	30:
		AssertTrue(Condition := rig.fbTel.bCloseRoofRequest, Message := 'latched after the hydraulics reset');
		F_Note(bFailed := NOT (rig.fbTel.bCloseRoofRequest), sText := CONCAT(sTest, 'latched after the hydraulics reset'));
		rig.fbTel.Reset();
		nStep := 40;
	40:
		AssertFalse(Condition := rig.fbTel.bCloseRoofRequest, Message := 'a reset without a cause clears it');
		F_Note(bFailed := (rig.fbTel.bCloseRoofRequest), sText := CONCAT(sTest, 'a reset without a cause clears it'));
		nStep := 99;
		TEST_FINISHED();
	END_CASE
END_IF
END_METHOD

// #24 step 7 PR 1 (D9, row E-stop): the E-stop sets bCloseRoofRequest. The E-stop circuit also cuts the roof drives, so the request
// must outlive it: a reset during the E-stop keeps it, it stays latched after the release, and only a reset without a cause
// clears it.
METHOD PRIVATE Roof_Request_On_Estop
VAR_INST
	rig			: FB_MonetRig;
	nStep		: INT;
	nCycles		: UINT;
	sTest		: STRING(80);
END_VAR
TEST('Roof_Request_On_Estop');
sTest := 'Roof_Request_On_Estop: ';
IF nStep >= 90 THEN
	RETURN;
END_IF
rig.Scan();
nCycles := nCycles + 1;
// one step every 3 scans: the cause or the reset of the step before has been scanned
IF nCycles >= 3 THEN
	nCycles := 0;
	CASE nStep OF
	0:
		AssertFalse(Condition := rig.fbTel.bCloseRoofRequest, Message := 'no request without a cause');
		F_Note(bFailed := (rig.fbTel.bCloseRoofRequest), sText := CONCAT(sTest, 'no request without a cause'));
		rig.SetEstop(TRUE);
		nStep := 10;
	10:
		AssertTrue(Condition := rig.fbTel.bCloseRoofRequest, Message := 'the E-stop sets the request');
		F_Note(bFailed := NOT (rig.fbTel.bCloseRoofRequest), sText := CONCAT(sTest, 'the E-stop sets the request'));
		rig.fbTel.Reset();
		nStep := 20;
	20:
		AssertTrue(Condition := rig.fbTel.bCloseRoofRequest, Message := 'a reset during the E-stop keeps it');
		F_Note(bFailed := NOT (rig.fbTel.bCloseRoofRequest), sText := CONCAT(sTest, 'a reset during the E-stop keeps it'));
		rig.SetEstop(FALSE);
		nStep := 30;
	30:
		AssertTrue(Condition := rig.fbTel.bCloseRoofRequest, Message := 'latched after the release');
		F_Note(bFailed := NOT (rig.fbTel.bCloseRoofRequest), sText := CONCAT(sTest, 'latched after the release'));
		// #24 step 7 PR 6: parked since the start, so the E-stop holds no park and nothing parks after the release
		AssertTrue(Condition := rig.fbTel.bIsParked AND NOT rig.fbTel.bParkActive AND rig.fbCovers.nCloseCalls = 0, Message := 'parked: no park after the release');
		F_Note(bFailed := NOT (rig.fbTel.bIsParked AND NOT rig.fbTel.bParkActive AND rig.fbCovers.nCloseCalls = 0), sText := CONCAT(sTest, 'parked: no park after the release'));
		rig.fbTel.Reset();
		nStep := 40;
	40:
		AssertFalse(Condition := rig.fbTel.bCloseRoofRequest, Message := 'a reset without a cause clears it');
		F_Note(bFailed := (rig.fbTel.bCloseRoofRequest), sText := CONCAT(sTest, 'a reset without a cause clears it'));
		nStep := 99;
		TEST_FINISHED();
	END_CASE
END_IF
END_METHOD

// #24 step 7 PR 1 (D9, row safety error): bSafetyError (SafetyHandling.error, no E-stop) sets bCloseRoofRequest; latched and reset
// as for the E-stop.
METHOD PRIVATE Roof_Request_On_Safety_Error
VAR_INST
	rig			: FB_MonetRig;
	nStep		: INT;
	nCycles		: UINT;
	sTest		: STRING(80);
END_VAR
TEST('Roof_Request_On_Safety_Error');
sTest := 'Roof_Request_On_Safety_Error: ';
IF nStep >= 90 THEN
	RETURN;
END_IF
rig.Scan();
nCycles := nCycles + 1;
// one step every 3 scans: the cause or the reset of the step before has been scanned
IF nCycles >= 3 THEN
	nCycles := 0;
	CASE nStep OF
	0:
		AssertFalse(Condition := rig.fbTel.bCloseRoofRequest, Message := 'no request without a cause');
		F_Note(bFailed := (rig.fbTel.bCloseRoofRequest), sText := CONCAT(sTest, 'no request without a cause'));
		rig.SetSafetyError(TRUE);
		nStep := 10;
	10:
		AssertTrue(Condition := rig.fbTel.bCloseRoofRequest, Message := 'the safety error sets the request');
		F_Note(bFailed := NOT (rig.fbTel.bCloseRoofRequest), sText := CONCAT(sTest, 'the safety error sets the request'));
		rig.fbTel.Reset();
		nStep := 20;
	20:
		AssertTrue(Condition := rig.fbTel.bCloseRoofRequest, Message := 'a reset with the safety error keeps it');
		F_Note(bFailed := NOT (rig.fbTel.bCloseRoofRequest), sText := CONCAT(sTest, 'a reset with the safety error keeps it'));
		rig.SetSafetyError(FALSE);
		nStep := 30;
	30:
		AssertTrue(Condition := rig.fbTel.bCloseRoofRequest, Message := 'latched after the safety error is gone');
		F_Note(bFailed := NOT (rig.fbTel.bCloseRoofRequest), sText := CONCAT(sTest, 'latched after the safety error is gone'));
		rig.fbTel.Reset();
		nStep := 40;
	40:
		AssertFalse(Condition := rig.fbTel.bCloseRoofRequest, Message := 'a reset without a cause clears it');
		F_Note(bFailed := (rig.fbTel.bCloseRoofRequest), sText := CONCAT(sTest, 'a reset without a cause clears it'));
		nStep := 99;
		TEST_FINISHED();
	END_CASE
END_IF
END_METHOD

// #24 step 7 PR 1 (D9, row power failure): bMainReady FALSE (PowerMonitoring.phaseOK) sets bCloseRoofRequest, so a phase dip that is
// gone again still requests the close; latched and reset as for the E-stop. Not M's bPowerFailure (a power-on failure).
METHOD PRIVATE Roof_Request_On_Power_Failure
VAR_INST
	rig			: FB_MonetRig;
	nStep		: INT;
	nCycles		: UINT;
	sTest		: STRING(80);
END_VAR
TEST('Roof_Request_On_Power_Failure');
sTest := 'Roof_Request_On_Power_Failure: ';
IF nStep >= 90 THEN
	RETURN;
END_IF
rig.Scan();
nCycles := nCycles + 1;
// one step every 3 scans: the cause or the reset of the step before has been scanned
IF nCycles >= 3 THEN
	nCycles := 0;
	CASE nStep OF
	0:
		AssertFalse(Condition := rig.fbTel.bCloseRoofRequest, Message := 'no request without a cause');
		F_Note(bFailed := (rig.fbTel.bCloseRoofRequest), sText := CONCAT(sTest, 'no request without a cause'));
		rig.SetMainReady(FALSE);
		nStep := 10;
	10:
		AssertTrue(Condition := rig.fbTel.bCloseRoofRequest, Message := 'the power failure sets the request');
		F_Note(bFailed := NOT (rig.fbTel.bCloseRoofRequest), sText := CONCAT(sTest, 'the power failure sets the request'));
		rig.fbTel.Reset();
		nStep := 20;
	20:
		AssertTrue(Condition := rig.fbTel.bCloseRoofRequest, Message := 'a reset during the power failure keeps it');
		F_Note(bFailed := NOT (rig.fbTel.bCloseRoofRequest), sText := CONCAT(sTest, 'a reset during the power failure keeps it'));
		rig.SetMainReady(TRUE);
		nStep := 30;
	30:
		AssertTrue(Condition := rig.fbTel.bCloseRoofRequest, Message := 'latched when the supply is back');
		F_Note(bFailed := NOT (rig.fbTel.bCloseRoofRequest), sText := CONCAT(sTest, 'latched when the supply is back'));
		rig.fbTel.Reset();
		nStep := 40;
	40:
		AssertFalse(Condition := rig.fbTel.bCloseRoofRequest, Message := 'a reset without a cause clears it');
		F_Note(bFailed := (rig.fbTel.bCloseRoofRequest), sText := CONCAT(sTest, 'a reset without a cause clears it'));
		nStep := 99;
		TEST_FINISHED();
	END_CASE
END_IF
END_METHOD

// #24 step 7 PR 1 (D9, row focus error): a focus error is a telescope error (bHwError, bError) but recoverable: no
// bCloseRoofRequest (open: plan 8.4). The software errors are checked in Goto_Times_Out_Ramps_Then_Drives_To_Park (16#10) and
// Invalid_Motion_Config_Is_Software_Error_32 (16#32).
METHOD PRIVATE No_Roof_Request_On_Focus_Error
VAR_INST
	rig			: FB_MonetRig;
	nStep		: INT;
	nCycles		: UINT;
	sTest		: STRING(80);
END_VAR
TEST('No_Roof_Request_On_Focus_Error');
sTest := 'No_Roof_Request_On_Focus_Error: ';
IF nStep >= 90 THEN
	RETURN;
END_IF
rig.Scan();
nCycles := nCycles + 1;
// one step every 3 scans: the cause or the reset of the step before has been scanned
IF nCycles >= 3 THEN
	nCycles := 0;
	CASE nStep OF
	0:
		rig.InjectFocusError(16#4550);
		nStep := 10;
	10:
		AssertTrue(Condition := rig.fbTel.bError, Message := 'the focus error is a telescope error');
		F_Note(bFailed := NOT (rig.fbTel.bError), sText := CONCAT(sTest, 'the focus error is a telescope error'));
		AssertFalse(Condition := rig.fbTel.bCloseRoofRequest, Message := 'no request for a focus error');
		F_Note(bFailed := (rig.fbTel.bCloseRoofRequest), sText := CONCAT(sTest, 'no request for a focus error'));
		nStep := 99;
		TEST_FINISHED();
	END_CASE
END_IF
END_METHOD

END_FUNCTION_BLOCK

(* stored: Version 1.1.0.1, ProductVersion 3.1.4024.15
   POU MonetSafeState_Tests: Id {d1a4e0f8-8062-4b9e-9210-d42d0064fb81}, SpecialFunc None
   Method Hydraulics_Error_While_Tracking_Ramps_Then_Parks_In_Place: Id {f533c953-e643-4316-8d3d-4e35919c0034}
   Method Hydraulics_Pressure_Loss_While_Tracking_Parks_In_Place_Without_Ramp: Id {c43e85dc-36d1-439d-a6ea-92bd15a671ca}
   Method Cover_Error_At_PowerOn_Fails_And_Stays_Parked: Id {916ea77f-2a49-49f8-8fa7-8ffe4aff53f2}
   Method Cover_Error_During_Park_Ends_The_Park_Without_Closed: Id {edc4f922-82f3-4352-b522-fd07dc3ed470}
   Method Cover_Error_While_Tracking_Drives_To_Park: Id {ce6d1ab5-6774-4afc-9d01-540fa1a2d1c3}
   Method Estop_During_Slew_Locks_Then_Parks_In_Place_After_The_Release: Id {8e60e5a2-3593-49f3-bb7c-2bde946b1ab4}
   Method Safety_Error_While_Tracking_Locks_Then_Parks_In_Place_When_It_Clears: Id {64191a98-fa3d-40d0-a9b1-c3c028f00663}
   Method Power_Failure_During_Goto_Ramps_Then_Parks_In_Place: Id {df52c504-416b-4fbe-ad2d-969ae710a1d6}
   Method Power_Failure_With_Pressure_Loss_Parks_In_Place_Without_Ramp: Id {c72128bf-20d1-403c-88a9-4a13e5bec2ac}
   Method Goto_Times_Out_Ramps_Then_Drives_To_Park: Id {575b45e8-d28e-4e1e-bc05-3296ec33c970}
   Method Home_Times_Out_Ramps_Then_Drives_To_Park: Id {452fcee1-58fd-44c6-bd2a-16a6b9438e2e}
   Method Clock_Invalid_Slew_Input_Is_Rejected: Id {3ae55bea-8d37-4402-9d1c-a6193ab6ddcb}
   Method Watchdog_Parks_And_Closes_The_Roof_In_One_Scan: Id {2ceca4cd-cb17-43a5-85a3-6b30784a4e38}
   Method Invalid_Motion_Config_Is_Software_Error_32: Id {1c5940e5-8f4f-45b6-867d-441dba951f47}
   Method Roof_Request_On_Axis_Errors: Id {7dd8bf42-fdcb-48ef-8970-6f1739a986dc}
   Method Roof_Request_On_Hydraulics_Error: Id {020b97fd-3bb6-4c6c-912e-b4e6b5eef17d}
   Method Roof_Request_On_Estop: Id {880f3c99-15e7-4f8e-8783-ead830e388fc}
   Method Roof_Request_On_Safety_Error: Id {81dfce06-d633-456d-ae15-e1171c532a06}
   Method Roof_Request_On_Power_Failure: Id {00264b16-ba15-4b5e-b428-f8b71d6b9d53}
   Method No_Roof_Request_On_Focus_Error: Id {750cde95-081b-44f0-9886-388f38ea3f96} *)
